(* IEC 61131-3 sources: Test-Git_ESME26/TestProgettoESME_26.fbsproj/AxisModuleLib Migration/AXM_FB_AxisModule.pou.xml.v3^, 40 files *)

(* ---- Additional_active.act.st ---- *)
__METADATA__
{
  "v3Meta": {
    "objectGuid": "95a41eea-732b-4df9-b4b6-dec268632541",
    "objectTypeGuid": "8ac092e5-3128-4e26-9e7e-11016c6684f2",
    "embeddedObjectTypeGuids": [
      "3b83b776-fb25-43b8-99f2-3c507c9143fc"
    ],
    "properties": {},
    "subObjects": {}
  }
}

iq_stAxisModuleItf.stMain.q_etOpMode := AXM_ET_OpMode.Additional;

xAdditionalStart := (xStartFlag OR iq_stAxisModuleItf.stMain.i_xStart) AND NOT stModuleReaction.axReaction[TPL.ET_Reaction.StopEndOfCycle];

iq_stAxisModuleItf.stAdditional.q_xEnable := xAdditionalEnable AND fbDriveEnable.q_xDriveEnabled;
iq_stAxisModuleItf.stAdditional.q_xStart := xAdditionalStart;
iq_stAxisModuleItf.stAdditional.q_xWsSelect := xWsSelect;
iq_stAxisModuleItf.stAdditional.q_xWsStart := xWsStartFlag;

IF iq_stAxisModuleItf.stAdditional.i_etDiag <> GD.ET_Diag.Ok THEN
	stExceptionModuleReaction2.etDiag := GD.ET_Diag.DiagActive;
	stExceptionModuleReaction2.udiDiagExt := AXM_ET_DiagExt.AdditionalModeException;
	stExceptionModuleReaction2.sMsg := SE_CTBX.FC_MultiConcat(	i_sString1 := GD.FC_EtDiagToString(i_etDiag := iq_stAxisModuleItf.stAdditional.i_etDiag),
															i_sString2 := ' ',
															i_sString3 := iq_stAxisModuleItf.stAdditional.i_sDiagExt,
															i_sString4 := SE_CTBX.FC_MultiConcat(	i_sString1 := '(',
																								i_sString2 := UDINT_TO_STRING(iq_stAxisModuleItf.stAdditional.i_udiDiagExt),
																								i_sString3 := ') ',
																								i_sString4 := iq_stAxisModuleItf.stAdditional.i_sMsg));
	ReportException(iq_stException := stExceptionModuleReaction2);
END_IF

xAdditionalActive := iq_stAxisModuleItf.stAdditional.i_xActive;

IF iq_stAxisModuleItf.stAdditional.i_xReady AND NOT iq_stAxisModuleItf.stAdditional.q_xStart THEN
	iq_stAxisModuleItf.stMain.q_etState := AXM_ET_State.AdditionalWaitForStart;
ELSIF iq_stAxisModuleItf.stAdditional.i_xReady AND iq_stAxisModuleItf.stAdditional.q_xStart THEN
	iq_stAxisModuleItf.stMain.q_etState := AXM_ET_State.AdditionalRunning;
ELSE
	IF xAdditionalEnable THEN
		iq_stAxisModuleItf.stMain.q_etState := AXM_ET_State.AdditionalInit;
	ELSE
		iq_stAxisModuleItf.stMain.q_etState := AXM_ET_State.AdditionalExit;
	END_IF
END_IF

(* ---- BrakeRelease_active.act.st ---- *)
__METADATA__
{
  "v3Meta": {
    "objectGuid": "62f6a697-2c31-4fa4-aead-e7013a7e303d",
    "objectTypeGuid": "8ac092e5-3128-4e26-9e7e-11016c6684f2",
    "embeddedObjectTypeGuids": [
      "3b83b776-fb25-43b8-99f2-3c507c9143fc"
    ],
    "properties": {},
    "subObjects": {}
  }
}

iq_stAxisModuleItf.stMain.q_etOpMode := AXM_ET_OpMode.BrakeRelease;

fbBrake(	i_xEnable			:= xBrakeEnable AND NOT fbDriveEnable.q_xDriveEnabled,
			i_xRelease			:= (xStartFlag OR iq_stAxisModuleItf.stMain.i_xStart),
			i_ifDrive			:= iq_stAxisModuleItf.stMain.i_ifDrive,
			q_xActive			=> ,
			q_xReady			=> ,
			q_xReleased			=> iq_stAxisModuleItf.stBrake.q_xBrakeReleased,
			q_etDiag			=> etDiagBuffer,
			q_etDiagExt			=> etDiagExtBufferPDL,
			q_sMsg				=> sDiagMsgBuffer);

DiagTestBrakeRelease(	iq_etDiag		:= fbBrake.q_etDiag,
						iq_etDiagExt	:= fbBrake.q_etDiagExt,
						iq_sMsg			:= fbBrake.q_sMsg);

IF fbBrake.q_xReady AND fbBrake.q_xReleased THEN
	iq_stAxisModuleItf.stMain.q_etState := AXM_ET_State.BrakeReleased;
ELSIF fbBrake.q_xReady AND NOT fbBrake.q_xReleased THEN
	iq_stAxisModuleItf.stMain.q_etState := AXM_ET_State.BrakeClosed;
ELSE
	IF xBrakeEnable THEN
		iq_stAxisModuleItf.stMain.q_etState := AXM_ET_State.BrakeReleaseInit;
	ELSE
		iq_stAxisModuleItf.stMain.q_etState := AXM_ET_State.BrakeReleaseExit;
	END_IF
END_IF

IF NOT xBrakeEnable AND NOT fbBrake.q_xActive THEN
	xBrakeActive := FALSE;
END_IF

(* ---- CancelException.meth.st ---- *)
{attribute 'conditionalshow_all_locals'}
METHOD INTERNAL CancelException
VAR_IN_OUT
	iq_stException	: TPL.ST_Exception;
END_VAR

TPL.FC_SetException(	i_xExceptionActive	:= FALSE,
						iq_stException		:= iq_stException,
						iq_stExceptionList	:= iq_stExceptionList,
						iq_stLogDataList	:= iq_stLogDataList,
						q_etDiag 			=> etDiagBuffer,
						q_etDiagExt 		=> etDiagExtBufferTPL,
						q_sMsg 				=> sDiagMsgBuffer);

(* ---- CheckCmd.meth.st ---- *)
{attribute 'conditionalshow_all_locals'}
METHOD INTERNAL CheckCmd
VAR_INPUT
END_VAR

(*--------------------------------------------------------------------------------------------------*)
(* CheckCMD is checking if CMD is supported by this module *)
(*--------------------------------------------------------------------------------------------------*)
xOpModeCmd:= FALSE;
xCheckCMDError:= FALSE;

IF iq_stStandardModuleItf.iq_diCmd = AXM_ET_Cmd.Homing OR
	iq_stStandardModuleItf.iq_diCmd = AXM_ET_Cmd.Manual OR
	iq_stStandardModuleItf.iq_diCmd = AXM_ET_Cmd.CamCs OR
	iq_stStandardModuleItf.iq_diCmd = AXM_ET_Cmd.CamWs OR
	iq_stStandardModuleItf.iq_diCmd = AXM_ET_Cmd.Endless OR
	iq_stStandardModuleItf.iq_diCmd = AXM_ET_Cmd.Positioning OR
	iq_stStandardModuleItf.iq_diCmd = AXM_ET_Cmd.BrakeRelease OR
	iq_stStandardModuleItf.iq_diCmd = AXM_ET_Cmd.AdditionalCs OR
	iq_stStandardModuleItf.iq_diCmd = AXM_ET_Cmd.AdditionalWs OR
	iq_stStandardModuleItf.iq_diCmd = AXM_ET_Cmd.DriveEnableOff OR
	iq_stStandardModuleItf.iq_diCmd = AXM_ET_Cmd.Stop THEN

	xOpModeCmd := TRUE;

ELSIF  iq_stStandardModuleItf.iq_diCmd = AXM_ET_Cmd.Start OR
		iq_stStandardModuleItf.iq_diCmd = AXM_ET_Cmd.StartTrig OR
		iq_stStandardModuleItf.iq_diCmd = AXM_ET_Cmd.StartTrigWaitInPos OR
		iq_stStandardModuleItf.iq_diCmd = AXM_ET_Cmd.Hold OR
		iq_stStandardModuleItf.iq_diCmd = AXM_ET_Cmd.WsStart OR
		iq_stStandardModuleItf.iq_diCmd = AXM_ET_Cmd.DriveEnableOn THEN

		xOpModeCmd:= FALSE;
ELSE
	xCheckCMDError := TRUE;
END_IF

(* ---- CmdControl_active.act.st ---- *)
__METADATA__
{
  "v3Meta": {
    "objectGuid": "07d6aa58-0565-4f47-8048-7bdd25741778",
    "objectTypeGuid": "8ac092e5-3128-4e26-9e7e-11016c6684f2",
    "embeddedObjectTypeGuids": [
      "3b83b776-fb25-43b8-99f2-3c507c9143fc"
    ],
    "properties": {},
    "subObjects": {}
  }
}

(* CMD execution

	algorithm:
	----------

	detect new command?
		check command?
			execute command;
		end
	end

	is command running (at least one cycle)?
		is command finished?
			signal success/unsuccessful
		end
	end
*)

xCommandAcceptedInThisCycle := FALSE;

(* Detect new command *)
IF(iq_stStandardModuleItf.i_xEnable) THEN
	IF (iq_stStandardModuleItf.iq_diCmd > 0 AND (NOT iq_stStandardModuleItf.q_xCmdActive (* In case no command is active *)
			OR iq_stStandardModuleItf.iq_diCmd <> iq_stStandardModuleItf.q_diCmdActive) (* In case a command is active *)) THEN

		xCommandRefused := FALSE; (* Flag is set by RefuseCommand() action *)

(****** Check if command execution is possible ******)
		CheckCMD();
		IF(xCheckCMDError) THEN
			(*** Check for unknown command ***)
			stExceptionCmdUnknown.sMsg := Standard.CONCAT('Cmd unknown: ',DINT_TO_STRING(iq_stStandardModuleItf.iq_diCmd));
			ReportException(iq_stException := stExceptionCmdUnknown);
			RefuseCommand();
		ELSE
			(*** Check for impossible overwrite ***)
			IF(iq_stStandardModuleItf.q_xCmdActive AND NOT((iq_stStandardModuleItf.iq_diCmd = AXM_ET_Cmd.Stop) OR
															(iq_stStandardModuleItf.iq_diCmd = AXM_ET_Cmd.BrakeRelease) OR
															((iq_stStandardModuleItf.iq_diCmd = AXM_ET_Cmd.Hold) AND (iq_stAxisModuleItf.stMain.q_etOpMode = AXM_ET_OpMode.Positioning) AND (iq_stStandardModuleItf.q_diCmdActive = AXM_ET_Cmd.Start)) OR
															((iq_stStandardModuleItf.iq_diCmd = AXM_ET_Cmd.Start) AND (iq_stAxisModuleItf.stMain.q_etOpMode = AXM_ET_OpMode.Endless) AND (iq_stStandardModuleItf.q_diCmdActive = AXM_ET_Cmd.Hold)))) THEN
				stExceptionCmdImpossibleOverwrite.sMsg := SE_CTBX.FC_MultiConcat(	i_sString1 := 'Cmd impossible: ',
																				//i_sString2 := iq_stStandardModuleItf.iq_diCmd
																				i_sString2 := AXM_FC_EtCmdToString(i_etCmd := iq_stStandardModuleItf.iq_diCmd),
																				i_sString3 := '; Cmd active: ',
																				i_sString4 := AXM_FC_EtCmdToString(i_etCmd := iq_stStandardModuleItf.q_diCmdActive) );
				ReportException(iq_stException := stExceptionCmdImpossibleOverwrite);
				RefuseCommand();
			ELSE
				(*** Check for impossible state ***)
				IF (((iq_stAxisModuleItf.stMain.q_etState = AXM_ET_State.NoOpDriveDisabled) OR (iq_stAxisModuleItf.stMain.q_etState = AXM_ET_State.NoOpDriveEnabled) ) AND
																								((iq_stStandardModuleItf.iq_diCmd = AXM_ET_Cmd.Start) OR
																								(iq_stStandardModuleItf.iq_diCmd = AXM_ET_Cmd.WsStart) OR
																								(iq_stStandardModuleItf.iq_diCmd = AXM_ET_Cmd.StartTrig) OR
																								(iq_stStandardModuleItf.iq_diCmd = AXM_ET_Cmd.StartTrigWaitInPos)) ) OR
					((iq_stAxisModuleItf.stMain.q_etState <> AXM_ET_State.MultiCamWaitForWsStart) AND (iq_stAxisModuleItf.stMain.q_etState <> AXM_ET_State.MultiCamRunning) AND (iq_stAxisModuleItf.stMain.q_etOpMode <> AXM_ET_OpMode.Additional) AND (iq_stStandardModuleItf.iq_diCmd = AXM_ET_Cmd.WsStart)) OR
					((iq_stAxisModuleItf.stMain.q_etState = AXM_ET_State.MultiCamWaitForWsStart) AND ((iq_stStandardModuleItf.iq_diCmd = AXM_ET_Cmd.WsStart) AND ((iq_stAxisModuleItf.stMultiCam.i_etWsMode = PDL_ET_MultiCamWsMode.StoredCamShowCamPosition) OR
																																		(iq_stAxisModuleItf.stMultiCam.i_etWsMode = PDL_ET_MultiCamWsMode.NewCamShowCamPosition)) ) ) OR
					((iq_stAxisModuleItf.stMain.q_etOpMode = AXM_ET_OpMode.Manual) AND ((iq_stStandardModuleItf.iq_diCmd = AXM_ET_Cmd.Hold) OR
																											(iq_stStandardModuleItf.iq_diCmd = AXM_ET_Cmd.Start)) ) OR
					((iq_stAxisModuleItf.stMain.q_etOpMode <> AXM_ET_OpMode.Positioning) AND (iq_stStandardModuleItf.iq_diCmd = AXM_ET_Cmd.StartTrigWaitInPos)) OR
					((iq_stAxisModuleItf.stMain.q_etOpMode <> AXM_ET_OpMode.Endless) AND (iq_stAxisModuleItf.stMain.q_etOpMode <> AXM_ET_OpMode.MultiCam) AND (iq_stAxisModuleItf.stMain.q_etOpMode <> AXM_ET_OpMode.Positioning) AND (iq_stStandardModuleItf.iq_diCmd = AXM_ET_Cmd.StartTrig))
					THEN
					stExceptionCmdImpossibleState.sMsg := SE_CTBX.FC_MultiConcat(	i_sString1 := 'Cmd impossible: ',
																				i_sString2 := AXM_FC_EtCmdToString(i_etCmd := iq_stStandardModuleItf.iq_diCmd),
																				i_sString3 := '; State: ',
																				i_sString4 := AXM_FC_EtStateToString(i_etState := iq_stAxisModuleItf.stMain.q_etState) );
					ReportException(iq_stException := stExceptionCmdImpossibleState);
					RefuseCommand();
				ELSIF ((iq_stAxisModuleItf.stMain.q_etOpMode = AXM_ET_OpMode.Homing OR
						iq_stAxisModuleItf.stMain.q_etOpMode = AXM_ET_OpMode.Manual OR
						iq_stAxisModuleItf.stMain.q_etOpMode = AXM_ET_OpMode.MultiCam OR
						iq_stAxisModuleItf.stMain.q_etOpMode = AXM_ET_OpMode.Endless OR
						iq_stAxisModuleItf.stMain.q_etOpMode = AXM_ET_OpMode.Positioning OR
						iq_stAxisModuleItf.stMain.q_etOpMode = AXM_ET_OpMode.BrakeRelease OR
						iq_stAxisModuleItf.stMain.q_etOpMode = AXM_ET_OpMode.Additional) AND ((iq_stAxisModuleItf.stMain.i_xStart OR xStartBitLastCycle) AND (iq_stStandardModuleItf.iq_diCMD = AXM_ET_Cmd.Start OR
																																						iq_stStandardModuleItf.iq_diCMD = AXM_ET_Cmd.Hold OR
																																						iq_stStandardModuleItf.iq_diCMD = AXM_ET_Cmd.StartTrig OR
																																						iq_stStandardModuleItf.iq_diCMD = AXM_ET_Cmd.StartTrigWaitInPos) )) THEN
					IF(iq_stAxisModuleItf.stMain.i_xStart) THEN
						stExceptionCmdImpossibleState.sMsg := SE_CTBX.FC_MultiConcat(	i_sString1 := 'Cmd impossible: ',
																					i_sString2 := AXM_FC_EtCmdToString(i_etCmd := iq_stStandardModuleItf.iq_diCmd),
																					i_sString3 := '; State: ',
																					i_sString4 := 'xStart input is TRUE');
						ReportException(iq_stException := stExceptionCmdImpossibleState);
						RefuseCommand();
					ELSE
						stExceptionCmdImpossibleState.sMsg := SE_CTBX.FC_MultiConcat(	i_sString1 := 'Cmd impossible: ',
																					i_sString2 := AXM_FC_EtCmdToString(i_etCmd := iq_stStandardModuleItf.iq_diCmd),
																					i_sString3 := '; State: ',
																					i_sString4 := 'xStart input was TRUE last cycle');
						ReportException(iq_stException := stExceptionCmdImpossibleState);
						RefuseCommand();
					END_IF
				ELSE
					(*** Check for impossible commands due to active error reactions ***)
					IF (stModuleReaction.axReaction[TPL.ET_Reaction.AsyncStop]
						OR stModuleReaction.axReaction[TPL.ET_Reaction.SyncStopEH]
						OR stModuleReaction.axReaction[TPL.ET_Reaction.SyncStopEL]
						OR stModuleReaction.axReaction[TPL.ET_Reaction.StopEndOfCycle])
						AND NOT (iq_stAxisModuleItf.stMain.q_etOpMode = AXM_ET_OpMode.BrakeRelease)
						AND	((iq_stStandardModuleItf.iq_diCmd = AXM_ET_Cmd.Start) OR
							(iq_stStandardModuleItf.iq_diCmd = AXM_ET_Cmd.WsStart) OR
							(iq_stStandardModuleItf.iq_diCmd = AXM_ET_Cmd.StartTrig) OR
							(iq_stStandardModuleItf.iq_diCmd = AXM_ET_Cmd.StartTrigWaitInPos)) THEN (* Start impossible if error reaction 4 or higher *)
							stWarningCmdImpossibleReaction.sMsg := SE_CTBX.FC_MultiConcat(	i_sString1 := 'Cmd impossible: ',
																						i_sString2 := AXM_FC_EtCmdToString(i_etCmd := iq_stStandardModuleItf.iq_diCmd),
																						i_sString3 := '; Reaction: ',
																						i_sString4 := TPL.FC_GetStandardReactionName(iq_stReaction := stModuleReaction));
							ReportException(iq_stException := stWarningCmdImpossibleReaction);
							RefuseCommand();
					ELSIF ((stModuleReaction.axReaction[TPL.ET_Reaction.AsyncStop]
							OR stModuleReaction.axReaction[TPL.ET_Reaction.SyncStopEH]
							OR stModuleReaction.axReaction[TPL.ET_Reaction.SyncStopEL] )
							AND xOpModeCmd AND
							NOT ((iq_stStandardModuleItf.iq_diCmd = AXM_ET_Cmd.Stop) OR (iq_stStandardModuleItf.iq_diCmd = AXM_ET_Cmd.DriveEnableOff) OR (iq_stStandardModuleItf.iq_diCmd = AXM_ET_Cmd.BrakeRelease)) ) THEN
							stWarningCmdImpossibleReaction.sMsg := SE_CTBX.FC_MultiConcat(	i_sString1 := 'Cmd impossible: ',
																						i_sString2 := AXM_FC_EtCmdToString(i_etCmd := iq_stStandardModuleItf.iq_diCmd),
																						i_sString3 := '; Reaction: ',
																						i_sString4 := TPL.FC_GetStandardReactionName(iq_stReaction := stModuleReaction));
							ReportException(iq_stException := stWarningCmdImpossibleReaction);
							RefuseCommand();
					ELSIF ((stModuleReaction.axReaction[TPL.ET_Reaction.AsyncStop]
							OR stModuleReaction.axReaction[TPL.ET_Reaction.SyncStopEL])
							AND (iq_stStandardModuleItf.iq_diCmd = AXM_ET_Cmd.DriveEnableOn)) THEN
							stWarningCmdImpossibleReaction.sMsg := SE_CTBX.FC_MultiConcat(	i_sString1 := 'Cmd impossible: ',
																						i_sString2 := AXM_FC_EtCmdToString(i_etCmd := iq_stStandardModuleItf.iq_diCmd),
																						i_sString3 := '; Reaction: ',
																						i_sString4 := TPL.FC_GetStandardReactionName(iq_stReaction := stModuleReaction));
							ReportException(iq_stException := stWarningCmdImpossibleReaction);
							RefuseCommand();
					END_IF
				END_IF
			END_IF
		END_IF

		IF(NOT xCommandRefused) THEN (* Command has passed all checks, execute command *)
			(* Accept command *)
			iq_stStandardModuleItf.q_xCmdActive := TRUE;
			iq_stStandardModuleItf.q_xCmdDone := FALSE;
			iq_stStandardModuleItf.q_diCmdActive := iq_stStandardModuleItf.iq_diCmd;

			xCommandAcceptedInThisCycle := TRUE; (* Signal for command done checks *)
			IF fbLoggerPoint.etLogLevel >= APL.ET_LogLevel.UserAction THEN
				fbLoggerPoint.AddLogEntry(	i_etLogLevel	:= APL.ET_LogLevel.UserAction,
											i_etDiag		:= GD.ET_Diag.Ok,
											i_udiDiagExt	:= AXM_ET_DiagExt.Ok,
											i_sMessage		:= Standard.CONCAT(Standard.CONCAT(Standard.CONCAT('Command executing: ', AXM_FC_EtCmdToString(i_etCmd := iq_stStandardModuleItf.iq_diCmd)),' number: '),DINT_TO_STRING(iq_stStandardModuleItf.iq_diCmd)),
											q_etDiag		:= ,
											q_etDiagExt		:= );
			END_IF

			IF(xOpModeCmd) THEN
				DisableAllJobs();
				xWsSelect			:= FALSE;
				xWsStartFlag		:= FALSE;

				CASE iq_stStandardModuleItf.iq_diCmd OF
				AXM_ET_Cmd.Stop:
					(* Do nothing, disabled OpMode flags automatically lead to NoOp *)
					xStartFlag := FALSE;

				AXM_ET_Cmd.Homing:
					xRefEnable := TRUE;

					IF iq_stAxisModuleItf.stHome.stSetPos.i_xKeepPowerDisabled AND
						( iq_stAxisModuleItf.stHome.i_etMode = PDL_ET_HomeMode.RestorePosFromAxisEncoder
						OR iq_stAxisModuleItf.stHome.i_etMode = PDL_ET_HomeMode.RestorePosFromRetain
						OR iq_stAxisModuleItf.stHome.i_etMode = PDL_ET_HomeMode.SetPosAxisAndLogEncoderPosition
						OR iq_stAxisModuleItf.stHome.i_etMode = PDL_ET_HomeMode.SetPosAxisPosition
						OR iq_stAxisModuleItf.stHome.i_etMode = PDL_ET_HomeMode.SetPosLogEncoderPosition )THEN
						xCMDPowerOn := FALSE;
					ELSE
						xCMDPowerOn := TRUE;
					END_IF

					IF NOT (iq_stAxisModuleItf.stMain.q_etOpMode = AXM_ET_OpMode.Homing) THEN
						xStartFlag := FALSE;
					END_IF

				AXM_ET_Cmd.Manual:
					xManEnable := TRUE;
					xCMDPowerOn := TRUE;

				AXM_ET_Cmd.CamCs:
					xCamEnable := TRUE;
					xCMDPowerOn := TRUE;
					xWsSelect := FALSE;
					xWsStartFlag := FALSE;
					IF NOT (iq_stAxisModuleItf.stMain.q_etOpMode = AXM_ET_OpMode.MultiCam) THEN
						xStartFlag := FALSE;
					END_IF

				AXM_ET_Cmd.CamWs:
					xCamEnable := TRUE;
					xCMDPowerOn := TRUE;
					xWsSelect := TRUE;
					xWsStartFlag := FALSE;
					IF NOT (iq_stAxisModuleItf.stMain.q_etOpMode = AXM_ET_OpMode.MultiCam) THEN
						xStartFlag := FALSE;
					END_IF

				AXM_ET_Cmd.Endless:
					xEndlessEnable := TRUE;
					xCMDPowerOn := TRUE;
					IF NOT (iq_stAxisModuleItf.stMain.q_etOpMode = AXM_ET_OpMode.Endless) THEN
						xStartFlag := FALSE;
					END_IF

				AXM_ET_Cmd.Positioning:
					xPosEnable := TRUE;
					xCMDPowerOn := TRUE;
					IF NOT (iq_stAxisModuleItf.stMain.q_etOpMode = AXM_ET_OpMode.Positioning) THEN
						xStartFlag := FALSE;
					END_IF

				AXM_ET_Cmd.BrakeRelease:
					xBrakeEnable := TRUE;
					xCMDPowerOn := FALSE;
					IF NOT (iq_stAxisModuleItf.stMain.q_etOpMode = AXM_ET_OpMode.BrakeRelease) THEN
						xStartFlag := FALSE;
					END_IF

				AXM_ET_Cmd.AdditionalCs:
					xAdditionalEnable := TRUE;
					xCMDPowerOn := TRUE;
					xWsSelect := FALSE;
					xWsStartFlag := FALSE;
					IF NOT (iq_stAxisModuleItf.stMain.q_etOpMode = AXM_ET_OpMode.Additional) THEN
						xStartFlag := FALSE;
					END_IF

				AXM_ET_Cmd.AdditionalWs:
					xAdditionalEnable := TRUE;
					xCMDPowerOn := TRUE;
					xWsSelect := TRUE;
					xWsStartFlag := FALSE;
					IF NOT (iq_stAxisModuleItf.stMain.q_etOpMode = AXM_ET_OpMode.Additional) THEN
						xStartFlag := FALSE;
					END_IF

				AXM_ET_Cmd.DriveEnableOff:
					xCMDPowerOn := FALSE;
					xStartFlag := FALSE;
				ELSE
					stExceptionModuleReaction1.etDiag := GD.ET_Diag.UnexpectedProgramBehavior;
					stExceptionModuleReaction1.udiDiagExt := AXM_ET_DiagExt.UnknownCase;
					stExceptionModuleReaction1.sMsg := '';
					ReportException(iq_stException := stExceptionModuleReaction1);
				END_CASE
			ELSE
				CASE iq_stStandardModuleItf.iq_diCmd OF
				AXM_ET_Cmd.Start:
					xStartFlag := TRUE;
					IF (iq_stAxisModuleItf.stMain.q_etOpMode = AXM_ET_OpMode.Homing) THEN
						(* Reset HomeOk when a new homing is started *)
						iq_stAxisModuleItf.stMain.q_xHomeOk := FALSE;
					END_IF

				AXM_ET_Cmd.StartTrig:
					xStartFlag := TRUE;

				AXM_ET_Cmd.StartTrigWaitInPos:
					xStartFlag := TRUE;

				AXM_ET_Cmd.WsStart:
					xWsStartFlag := TRUE;
					(* In additional mode it has to be possible to set WsStart independent of start *)
					IF NOT (iq_stAxisModuleItf.stMain.q_etOpMode = AXM_ET_OpMode.Additional) THEN
						xStartFlag  := TRUE;
					END_IF

				AXM_ET_Cmd.Hold:
					xStartFlag := FALSE;

				AXM_ET_Cmd.DriveEnableOn:
					xCMDPowerOn := TRUE;

				ELSE
					stExceptionModuleReaction1.etDiag := GD.ET_Diag.UnexpectedProgramBehavior;
					stExceptionModuleReaction1.udiDiagExt := AXM_ET_DiagExt.UnknownCase;
					stExceptionModuleReaction1.sMsg := '';
					ReportException(iq_stException := stExceptionModuleReaction1);
				END_CASE

			END_IF
		END_IF (* New command? *)
	END_IF

(********************************************* Check successful and unsucessful of given commands ****************************************)

	(* Check if active command is done or is stopped by an error *)
	IF(NOT xCommandAcceptedInThisCycle) THEN (* Don't execute these checks if we accepted a new command in this cycle
		to ensure that execution of every command requires a minimum of 2 cycles *)

		IF(iq_stStandardModuleItf.q_xCmdActive) THEN
			CASE iq_stStandardModuleItf.iq_diCmd OF
			AXM_ET_Cmd.Homing:
				(* Successful *)
				IF (iq_stAxisModuleItf.stMain.q_etOpMode = AXM_ET_OpMode.Homing) AND NOT (iq_stAxisModuleItf.stMain.q_etState = AXM_ET_State.HomingInit) THEN
					SignalSuccessfulExecution();
				END_IF
				(* Unsucessful *)
				IF(stModuleReaction.axReaction[TPL.ET_Reaction.AsyncStop]
					OR stModuleReaction.axReaction[TPL.ET_Reaction.SyncStopEH]
					OR stModuleReaction.axReaction[TPL.ET_Reaction.SyncStopEL]) THEN
					SignalUnsuccessfulExecution();
				END_IF

			AXM_ET_Cmd.Manual:
				(* Successful *)
				IF (iq_stAxisModuleItf.stMain.q_etOpMode = AXM_ET_OpMode.Manual) AND NOT (iq_stAxisModuleItf.stMain.q_etState = AXM_ET_State.ManualInit) THEN
					SignalSuccessfulExecution();
				END_IF
				(* Unsucessful *)
				IF(stModuleReaction.axReaction[TPL.ET_Reaction.AsyncStop]
					OR stModuleReaction.axReaction[TPL.ET_Reaction.SyncStopEH]
					OR stModuleReaction.axReaction[TPL.ET_Reaction.SyncStopEL]) THEN
					SignalUnsuccessfulExecution();
				END_IF

			AXM_ET_Cmd.CamCs:
				(* Successful *)
				IF (iq_stAxisModuleItf.stMain.q_etOpMode = AXM_ET_OpMode.MultiCam) AND NOT (iq_stAxisModuleItf.stMain.q_etState = AXM_ET_State.MultiCamInit) THEN
					SignalSuccessfulExecution();
				END_IF
				(* Unsucessful *)
				IF(stModuleReaction.axReaction[TPL.ET_Reaction.AsyncStop]
					OR stModuleReaction.axReaction[TPL.ET_Reaction.SyncStopEH]
					OR stModuleReaction.axReaction[TPL.ET_Reaction.SyncStopEL]) THEN
					SignalUnsuccessfulExecution();
				END_IF

			AXM_ET_Cmd.CamWs:
				(* Successful *)
				IF (iq_stAxisModuleItf.stMain.q_etOpMode = AXM_ET_OpMode.MultiCam) AND NOT (iq_stAxisModuleItf.stMain.q_etState = AXM_ET_State.MultiCamInit) THEN
					SignalSuccessfulExecution();
				END_IF
				(* Unsucessful *)
				IF(stModuleReaction.axReaction[TPL.ET_Reaction.AsyncStop]
					OR stModuleReaction.axReaction[TPL.ET_Reaction.SyncStopEH]
					OR stModuleReaction.axReaction[TPL.ET_Reaction.SyncStopEL]) THEN
					SignalUnsuccessfulExecution();
				END_IF

			AXM_ET_Cmd.Endless:
				(* Successful *)
				IF (iq_stAxisModuleItf.stMain.q_etOpMode = AXM_ET_OpMode.Endless) AND NOT (iq_stAxisModuleItf.stMain.q_etState = AXM_ET_State.EndlessInit) THEN
					SignalSuccessfulExecution();
				END_IF
				(* Unsucessful *)
				IF(stModuleReaction.axReaction[TPL.ET_Reaction.AsyncStop]
					OR stModuleReaction.axReaction[TPL.ET_Reaction.SyncStopEH]
					OR stModuleReaction.axReaction[TPL.ET_Reaction.SyncStopEL]) THEN
					SignalUnsuccessfulExecution();
				END_IF

			AXM_ET_Cmd.Positioning:
				(* Successful *)
				IF (iq_stAxisModuleItf.stMain.q_etOpMode = AXM_ET_OpMode.Positioning) AND NOT (iq_stAxisModuleItf.stMain.q_etState = AXM_ET_State.PositioningInit) THEN
					SignalSuccessfulExecution();
				END_IF
				(* Unsucessful *)
				IF(stModuleReaction.axReaction[TPL.ET_Reaction.AsyncStop]
					OR stModuleReaction.axReaction[TPL.ET_Reaction.SyncStopEH]
					OR stModuleReaction.axReaction[TPL.ET_Reaction.SyncStopEL]) THEN
					SignalUnsuccessfulExecution();
				END_IF

			AXM_ET_Cmd.BrakeRelease:
				(* Successful *)
				IF (iq_stAxisModuleItf.stMain.q_etOpMode = AXM_ET_OpMode.BrakeRelease) AND
					( (NOT fbBrake.i_xRelease AND (iq_stAxisModuleItf.stMain.q_etState = AXM_ET_State.BrakeClosed)) OR
					(fbBrake.i_xRelease AND (iq_stAxisModuleItf.stMain.q_etState = AXM_ET_State.BrakeReleased)) ) THEN
					// real axis can still be in state brake open if gone to brake release opmode,
					// therefore delay signal cmd successfull till brake closed is reached
					SignalSuccessfulExecution();
				END_IF

			AXM_ET_Cmd.AdditionalCs:
				(* Successful *)
				IF (iq_stAxisModuleItf.stMain.q_etOpMode = AXM_ET_OpMode.Additional) AND NOT (iq_stAxisModuleItf.stMain.q_etState = AXM_ET_State.AdditionalInit) THEN
					SignalSuccessfulExecution();
				END_IF
				(* Unsucessful *)
				IF(stModuleReaction.axReaction[TPL.ET_Reaction.AsyncStop]
					OR stModuleReaction.axReaction[TPL.ET_Reaction.SyncStopEH]
					OR stModuleReaction.axReaction[TPL.ET_Reaction.SyncStopEL]) THEN
					SignalUnsuccessfulExecution();
				END_IF

			AXM_ET_Cmd.AdditionalWs:
				(* Successful *)
				IF (iq_stAxisModuleItf.stMain.q_etOpMode = AXM_ET_OpMode.Additional) AND NOT (iq_stAxisModuleItf.stMain.q_etState = AXM_ET_State.AdditionalInit) THEN
					SignalSuccessfulExecution();
				END_IF
				(* Unsucessful *)
				IF(stModuleReaction.axReaction[TPL.ET_Reaction.AsyncStop]
					OR stModuleReaction.axReaction[TPL.ET_Reaction.SyncStopEH]
					OR stModuleReaction.axReaction[TPL.ET_Reaction.SyncStopEL]) THEN
					SignalUnsuccessfulExecution();
				END_IF

			AXM_ET_Cmd.Start:
				(* Successful *)
				IF ((iq_stAxisModuleItf.stMain.q_etState = AXM_ET_State.HomingWaitForStart) AND iq_stAxisModuleItf.stMain.q_xHomeOk) OR
					(iq_stAxisModuleItf.stMain.q_etState = AXM_ET_State.HomingDone) OR
					(iq_stAxisModuleItf.stMain.q_etState = AXM_ET_State.MultiCamWaitForWsStart) OR
					(iq_stAxisModuleItf.stMain.q_etState = AXM_ET_State.MultiCamRunning) OR
					(iq_stAxisModuleItf.stMain.q_etState = AXM_ET_State.EndlessRunning) OR
					(iq_stAxisModuleItf.stMain.q_etState = AXM_ET_State.PositioningRunning) OR
					(iq_stAxisModuleItf.stMain.q_etState = AXM_ET_State.BrakeReleased) OR
					((iq_stAxisModuleItf.stMain.q_etOpMode = AXM_ET_OpMode.Additional) AND iq_stAxisModuleItf.stAdditional.i_xActionCmdDone) THEN
					SignalSuccessfulExecution();
				END_IF
				(* Unsucesful *)
				IF(stModuleReaction.axReaction[TPL.ET_Reaction.AsyncStop]
					OR stModuleReaction.axReaction[TPL.ET_Reaction.SyncStopEH]
					OR stModuleReaction.axReaction[TPL.ET_Reaction.SyncStopEL]
					OR stModuleReaction.axReaction[TPL.ET_Reaction.StopEndOfCycle])
					AND NOT (iq_stAxisModuleItf.stMain.q_etOpMode = AXM_ET_OpMode.BrakeRelease) THEN
					SignalUnsuccessfulExecution();
				END_IF

			AXM_ET_Cmd.StartTrig:
				(* Successful *)
				IF (iq_stAxisModuleItf.stMain.q_etState = AXM_ET_State.PositioningRunning) OR
					(iq_stAxisModuleItf.stMain.q_etState = AXM_ET_State.MultiCamRunning) OR
					(iq_stAxisModuleItf.stMain.q_etState = AXM_ET_State.EndlessRunning) THEN
					xStartFlag := FALSE;
					SignalSuccessfulExecution();
				END_IF
				(* Unsucesful *)
				IF(stModuleReaction.axReaction[TPL.ET_Reaction.AsyncStop]
					OR stModuleReaction.axReaction[TPL.ET_Reaction.SyncStopEH]
					OR stModuleReaction.axReaction[TPL.ET_Reaction.SyncStopEL]
					)
					AND NOT (iq_stAxisModuleItf.stMain.q_etOpMode = AXM_ET_OpMode.BrakeRelease) THEN
					SignalUnsuccessfulExecution();
				END_IF

			AXM_ET_Cmd.StartTrigWaitInPos:
				(* Successful *)
				IF fbVarioPos.q_xInPosition THEN
					xStartFlag := FALSE;
					SignalSuccessfulExecution();
				END_IF
				(* Unsucesful *)
				IF(stModuleReaction.axReaction[TPL.ET_Reaction.AsyncStop]
					OR stModuleReaction.axReaction[TPL.ET_Reaction.SyncStopEH]
					OR stModuleReaction.axReaction[TPL.ET_Reaction.SyncStopEL]
					)
					AND NOT (iq_stAxisModuleItf.stMain.q_etOpMode = AXM_ET_OpMode.BrakeRelease) THEN
					SignalUnsuccessfulExecution();
				END_IF

			AXM_ET_Cmd.Stop:
				(* Successful *)
				IF (iq_stAxisModuleItf.stMain.q_etState = AXM_ET_State.NoOpDriveDisabled) OR
					(iq_stAxisModuleItf.stMain.q_etState = AXM_ET_State.NoOpDriveEnabled) THEN
					iq_stAxisModuleItf.stMain.q_etOpMode := AXM_ET_OpMode.NoOp;
					SignalSuccessfulExecution();
				END_IF

			AXM_ET_Cmd.Hold:
				IF iq_stAxisModuleItf.stMain.i_xStart THEN
					stExceptionModuleReaction2.sMsg := 'rising edge of xStart input during execution of CMD Hold';
					ReportException(iq_stException := stExceptionModuleReaction2);
					RefuseCommand();
				ELSIF (* Successful *)
					(iq_stAxisModuleItf.stMain.q_etState = AXM_ET_State.HomingWaitForStart) OR
					(iq_stAxisModuleItf.stMain.q_etState = AXM_ET_State.MultiCamWaitForStart) OR
					(iq_stAxisModuleItf.stMain.q_etState = AXM_ET_State.EndlessWaitForStart) OR
					(iq_stAxisModuleItf.stMain.q_etState = AXM_ET_State.PositioningWaitForStart) OR
					(iq_stAxisModuleItf.stMain.q_etState = AXM_ET_State.BrakeClosed) OR
					(iq_stAxisModuleItf.stMain.q_etState = AXM_ET_State.AdditionalWaitForStart) OR
					(iq_stAxisModuleItf.stMain.q_etState = AXM_ET_State.NoOpDriveDisabled) OR
					(iq_stAxisModuleItf.stMain.q_etState = AXM_ET_State.NoOpDriveEnabled) OR
					((iq_stAxisModuleItf.stMain.q_etOpMode = AXM_ET_OpMode.Additional) AND iq_stAxisModuleItf.stAdditional.i_xActionCmdDone) THEN
					SignalSuccessfulExecution();
				ELSIF (* Unsucessful *)
					(stModuleReaction.axReaction[TPL.ET_Reaction.AsyncStop]
					OR stModuleReaction.axReaction[TPL.ET_Reaction.SyncStopEH]
					OR stModuleReaction.axReaction[TPL.ET_Reaction.SyncStopEL]) AND NOT (iq_stAxisModuleItf.stMain.q_etOpMode = AXM_ET_OpMode.BrakeRelease) THEN
					SignalUnsuccessfulExecution();
				END_IF

			AXM_ET_Cmd.WsStart:
				(* Successful *)
				IF ((iq_stAxisModuleItf.stMain.q_etState = AXM_ET_State.HomingWaitForStart) AND iq_stAxisModuleItf.stMain.q_xHomeOk) OR
					(iq_stAxisModuleItf.stMain.q_etState = AXM_ET_State.MultiCamRunning) OR
					(iq_stAxisModuleItf.stMain.q_etState = AXM_ET_State.EndlessRunning) OR
					(iq_stAxisModuleItf.stMain.q_etState = AXM_ET_State.PositioningRunning) OR
					(iq_stAxisModuleItf.stMain.q_etState = AXM_ET_State.BrakeReleased) OR
					((iq_stAxisModuleItf.stMain.q_etOpMode = AXM_ET_OpMode.Additional) AND iq_stAxisModuleItf.stAdditional.i_xActionCmdDone) THEN
					SignalSuccessfulExecution();
				END_IF
				(* Unsucesful *)
				IF(stModuleReaction.axReaction[TPL.ET_Reaction.AsyncStop]
					OR stModuleReaction.axReaction[TPL.ET_Reaction.SyncStopEH]
					OR stModuleReaction.axReaction[TPL.ET_Reaction.SyncStopEL]
					OR stModuleReaction.axReaction[TPL.ET_Reaction.StopEndOfCycle]) THEN
					SignalUnsuccessfulExecution();
				END_IF

			AXM_ET_Cmd.DriveEnableOn:
				(* Successful *)
				IF(etPowerState = AXM_ET_PowerState.PowerOn) THEN
					SignalSuccessfulExecution();
				END_IF
				(* Unsucessful *)
				IF(stModuleReaction.axReaction[TPL.ET_Reaction.AsyncStop]
					OR stModuleReaction.axReaction[TPL.ET_Reaction.SyncStopEH]
					OR stModuleReaction.axReaction[TPL.ET_Reaction.SyncStopEL]) THEN
					SignalUnsuccessfulExecution();
				END_IF

			AXM_ET_Cmd.DriveEnableOff:
				(* Successful *)
				IF(etPowerState = AXM_ET_PowerState.PowerOff) THEN
					SignalSuccessfulExecution();
				END_IF

			ELSE
				stExceptionModuleReaction1.etDiag := GD.ET_Diag.UnexpectedProgramBehavior;
				stExceptionModuleReaction1.udiDiagExt := AXM_ET_DiagExt.UnknownCase;
				stExceptionModuleReaction1.sMsg := '';
				ReportException(iq_stException := stExceptionModuleReaction1);
			END_CASE
		END_IF
	END_IF
ELSE
	(* Module is going to be disabled *)
	IF xEnableFlag THEN
		etPowerState := AXM_ET_PowerState.WaitForDisabled;
		IF fbLoggerPoint.etLogLevel >= APL.ET_LogLevel.UserAction THEN
			fbLoggerPoint.AddLogEntry(	i_etLogLevel	:= APL.ET_LogLevel.UserAction,
										i_etDiag		:= GD.ET_Diag.Ok,
										i_udiDiagExt	:= AXM_ET_DiagExt.Ok,
										i_sMessage		:= 'disabeling Module',
										q_etDiag		:= ,
										q_etDiagExt		:= );
		END_IF
	END_IF
	iq_stStandardModuleItf.q_xReady := FALSE;
	xEnableFlag := FALSE;
	xCMDPowerOn := FALSE;
	DisableAllJobs();
	xStartFlag := FALSE;
	xWsSelect := FALSE;
	xWsStartFlag := FALSE;
	IF(iq_stStandardModuleItf.q_xCmdActive) THEN (* If a command is currently active, cancel its execution *)
		SignalUnsuccessfulExecution();
	ELSE
		InactiveCmdExecution(); (* Command processing as if we were disabled *)
	END_IF
END_IF
xStartBitLastCycle := iq_stAxisModuleItf.stMain.i_xStart;

(* ---- DiagQuit.meth.st ---- *)
{attribute 'conditionalshow_all_locals'}
METHOD INTERNAL DiagQuit
VAR_INPUT
END_VAR

IF(iq_stStandardModuleItf.i_xDiagQuit AND NOT xDiagQuitFlag) THEN
	(* Rising edge of error quit *)
	xDiagQuitFlag := TRUE;
	xNotAbleToSetException := FALSE;
	iq_stStandardModuleItf.q_xException := FALSE;

	FOR udii := 1 TO TPL.ET_Reaction.MainsContactorOff DO
		stLocalReaction.axReaction[udii] := FALSE;
	END_FOR

	IF(iq_stStandardModuleItf.iq_diCMD < 0) THEN
		iq_stStandardModuleItf.iq_diCMD := 0;
	END_IF
	IF fbLoggerPoint.etLogLevel >= APL.ET_LogLevel.UserAction THEN
		fbLoggerPoint.AddLogEntry(	i_etLogLevel	:= APL.ET_LogLevel.UserAction,
									i_etDiag		:= GD.ET_Diag.Ok,
									i_udiDiagExt	:= AXM_ET_DiagExt.Ok,
									i_sMessage		:= 'Diag Quit',
									q_etDiag		:= ,
									q_etDiagExt		:= );
	END_IF
ELSIF(NOT iq_stStandardModuleItf.i_xDiagQuit AND xDiagQuitFlag) THEN
	xDiagQuitFlag := FALSE;
END_IF

(* ---- DiagTestBrakeRelease.meth.st ---- *)
{attribute 'conditionalshow_all_locals'}
METHOD INTERNAL DiagTestBrakeRelease
VAR_IN_OUT
	iq_etDiag		: GD.ET_Diag;
	iq_etDiagExt	: PDL_ET_DiagExt;
	iq_sMsg			: STRING[80];
END_VAR

IF (iq_etDiag <> GD.ET_Diag.Ok) THEN
	CASE iq_etDiagExt OF

	PDL_ET_DiagExt.DriveInvalid: (* if Drive has no brake *)
		stExceptionModuleReaction2.etDiag := GD.ET_Diag.InputParameterInvalid;
		stExceptionModuleReaction2.udiDiagExt := AXM_ET_DiagExt.DriveInvalid;
		stExceptionModuleReaction2.sMsg := iq_sMsg;
		ReportException(iq_stException := stExceptionModuleReaction2);

	PDL_ET_DiagExt.DriveNotReady:
		stExceptionModuleReaction2.etDiag := GD.ET_Diag.DriveConditionInvalid;
		stExceptionModuleReaction2.udiDiagExt := AXM_ET_DiagExt.DriveNotReady;
		stExceptionModuleReaction2.sMsg := iq_sMsg;
		ReportException(iq_stException := stExceptionModuleReaction2);

	ELSE
		stExceptionUnexpected.udiDiagExt := AXM_ET_DiagExt.UnexpectedFeedback;
		stExceptionUnexpected.sMsg := SE_CTBX.FC_MultiConcat(	i_sString1 := 'FB_BrakeRelease ',
															i_sString2 := PDL_FC_EtDiagExtToString(i_etDiagExt := iq_etDiagExt),
															i_sString3 := ' ',
															i_sString4 := iq_sMsg);
		ReportException(iq_stException := stExceptionUnexpected);
	END_CASE
END_IF

(* ---- DiagTestDriveEnable.meth.st ---- *)
{attribute 'conditionalshow_all_locals'}
METHOD INTERNAL DiagTestDriveEnable
VAR_IN_OUT
	iq_etDiag		: GD.ET_Diag;
	iq_etDiagExt	: PDL_ET_DiagExt;
	iq_sMsg			: STRING[80];
END_VAR

IF (iq_etDiag <> GD.ET_Diag.Ok) THEN
	CASE iq_etDiagExt OF
	PDL_ET_DiagExt.DriveNotReady:
		stExceptionModuleReaction2.etDiag := GD.ET_Diag.DriveConditionInvalid;
		stExceptionModuleReaction2.udiDiagExt := AXM_ET_DiagExt.DriveNotReady;
		stExceptionModuleReaction2.sMsg := iq_sMsg;
		ReportException(iq_stException := stExceptionModuleReaction2);

	PDL_ET_DiagExt.InverterEnableOff:
		stExceptionModuleReaction2.etDiag := GD.ET_Diag.DriveConditionInvalid;
		stExceptionModuleReaction2.udiDiagExt := AXM_ET_DiagExt.InverterEnableOff;
		stExceptionModuleReaction2.sMsg := iq_sMsg;
		ReportException(iq_stException := stExceptionModuleReaction2);

	PDL_ET_DiagExt.TorqueEnableOff:
		stExceptionModuleReaction2.etDiag := GD.ET_Diag.DriveConditionInvalid;
		stExceptionModuleReaction2.udiDiagExt := AXM_ET_DiagExt.TorqueEnableOff;
		stExceptionModuleReaction2.sMsg := iq_sMsg;
		ReportException(iq_stException := stExceptionModuleReaction2);

	PDL_ET_DiagExt.PowerSupplyInvalid:
		stExceptionModuleReaction2.etDiag := GD.ET_Diag.InputParameterInvalid;
		stExceptionModuleReaction2.udiDiagExt := AXM_ET_DiagExt.PowerSupplyInvalid;
		stExceptionModuleReaction2.sMsg := iq_sMsg;
		ReportException(iq_stException := stExceptionModuleReaction2);

	PDL_ET_DiagExt.PowerSupplyNotFound:
		stExceptionModuleReaction2.etDiag := GD.ET_Diag.InputParameterInvalid;
		stExceptionModuleReaction2.udiDiagExt := AXM_ET_DiagExt.PowerSupplyNotFound;
		stExceptionModuleReaction2.sMsg := iq_sMsg;
		ReportException(iq_stException := stExceptionModuleReaction2);

	PDL_ET_DiagExt.PowerSupplyNotReady:
		stExceptionModuleReaction2.etDiag := GD.ET_Diag.PowerSupplyConditionInvalid;
		stExceptionModuleReaction2.udiDiagExt := AXM_ET_DiagExt.PowerSupplyNotReady;
		stExceptionModuleReaction2.sMsg := iq_sMsg;
		ReportException(iq_stException := stExceptionModuleReaction2);

	ELSE
		stExceptionUnexpected.udiDiagExt := AXM_ET_DiagExt.UnexpectedFeedback;
		stExceptionUnexpected.sMsg := SE_CTBX.FC_MultiConcat(	i_sString1 := 'FB_DriveEnable ',
															i_sString2 := PDL_FC_EtDiagExtToString(i_etDiagExt := iq_etDiagExt),
															i_sString3 := ' ',
															i_sString4 := iq_sMsg);
		ReportException(iq_stException := stExceptionUnexpected);
	END_CASE
END_IF

(* ---- DiagTestEndless.meth.st ---- *)
{attribute 'conditionalshow_all_locals'}
METHOD INTERNAL DiagTestEndless
VAR_IN_OUT
	iq_etDiag		: GD.ET_Diag;
	iq_etDiagExt	: PDL_ET_DiagExt;
	iq_sMsg			: STRING[80];
END_VAR

IF (iq_etDiag <> GD.ET_Diag.Ok) THEN
	CASE iq_etDiagExt OF
	PDL_ET_DiagExt.VelRange:
		stExceptionModuleReaction2.etDiag := GD.ET_Diag.InputParameterInvalid;
		stExceptionModuleReaction2.udiDiagExt := AXM_ET_DiagExt.VelRange;
		stExceptionModuleReaction2.sMsg := iq_sMsg;
		ReportException(iq_stException := stExceptionModuleReaction2);

	PDL_ET_DiagExt.AccRange:
		stExceptionModuleReaction2.etDiag := GD.ET_Diag.InputParameterInvalid;
		stExceptionModuleReaction2.udiDiagExt := AXM_ET_DiagExt.AccRange;
		stExceptionModuleReaction2.sMsg := iq_sMsg;
		ReportException(iq_stException := stExceptionModuleReaction2);

	PDL_ET_DiagExt.DecRange:
		stExceptionModuleReaction2.etDiag := GD.ET_Diag.InputParameterInvalid;
		stExceptionModuleReaction2.udiDiagExt := AXM_ET_DiagExt.DecRange;
		stExceptionModuleReaction2.sMsg := iq_sMsg;
		ReportException(iq_stException := stExceptionModuleReaction2);

	PDL_ET_DiagExt.JerkRange:
		stExceptionModuleReaction2.etDiag := GD.ET_Diag.InputParameterInvalid;
		stExceptionModuleReaction2.udiDiagExt := AXM_ET_DiagExt.JerkRange;
		stExceptionModuleReaction2.sMsg := iq_sMsg;
		ReportException(iq_stException := stExceptionModuleReaction2);

	PDL_ET_DiagExt.PeriodRange:
		stExceptionModuleReaction2.etDiag := GD.ET_Diag.InputParameterInvalid;
		stExceptionModuleReaction2.udiDiagExt := AXM_ET_DiagExt.PeriodRange;
		stExceptionModuleReaction2.sMsg := iq_sMsg;
		ReportException(iq_stException := stExceptionModuleReaction2);

	PDL_ET_DiagExt.StopPositionRange:
		stExceptionModuleReaction2.etDiag := GD.ET_Diag.InputParameterInvalid;
		stExceptionModuleReaction2.udiDiagExt := AXM_ET_DiagExt.StopPositionRange;
		stExceptionModuleReaction2.sMsg := iq_sMsg;
		ReportException(iq_stException := stExceptionModuleReaction2);

	ELSE
		stExceptionUnexpected.udiDiagExt := AXM_ET_DiagExt.UnexpectedFeedback;
		stExceptionUnexpected.sMsg := SE_CTBX.FC_MultiConcat(	i_sString1 := 'FB_Endless ',
															i_sString2 := PDL_FC_EtDiagExtToString(i_etDiagExt := iq_etDiagExt),
															i_sString3 := ' ',
															i_sString4 := iq_sMsg);
		ReportException(iq_stException := stExceptionUnexpected);
	END_CASE
END_IF

(* ---- DiagTestHoming.meth.st ---- *)
{attribute 'conditionalshow_all_locals'}
METHOD INTERNAL DiagTestHoming
VAR_IN_OUT
	iq_etDiag		: GD.ET_Diag;
	iq_etDiagExt	: PDL_ET_DiagExt;
	iq_sMsg			: STRING[80];
END_VAR

IF (iq_etDiag <> GD.ET_Diag.Ok) THEN
	CASE iq_etDiagExt OF
	PDL_ET_DiagExt.AbsEncOffsetRange:
		stExceptionModuleReaction2.etDiag := GD.ET_Diag.InputParameterInvalid;
		stExceptionModuleReaction2.udiDiagExt := AXM_ET_DiagExt.AbsEncOffsetRange;
		stExceptionModuleReaction2.sMsg := iq_sMsg;
		ReportException(iq_stException := stExceptionModuleReaction2);

	PDL_ET_DiagExt.AccRange:
		stExceptionModuleReaction2.etDiag := GD.ET_Diag.InputParameterInvalid;
		stExceptionModuleReaction2.udiDiagExt := AXM_ET_DiagExt.AccRange;
		stExceptionModuleReaction2.sMsg := iq_sMsg;
		ReportException(iq_stException := stExceptionModuleReaction2);

	PDL_ET_DiagExt.CheckSumInvalid:
		stExceptionModuleReaction2.etDiag := GD.ET_Diag.InputParameterInvalid;
		stExceptionModuleReaction2.udiDiagExt := AXM_ET_DiagExt.CheckSumInvalid;
		stExceptionModuleReaction2.sMsg := iq_sMsg;
		ReportException(iq_stException := stExceptionModuleReaction2);

	PDL_ET_DiagExt.DataNVRamInvalid:
		stExceptionModuleReaction2.etDiag := GD.ET_Diag.InputParameterInvalid;
		stExceptionModuleReaction2.udiDiagExt := AXM_ET_DiagExt.DataNVRamInvalid;
		stExceptionModuleReaction2.sMsg := iq_sMsg;
		ReportException(iq_stException := stExceptionModuleReaction2);

	PDL_ET_DiagExt.DecRange:
		stExceptionModuleReaction2.etDiag := GD.ET_Diag.InputParameterInvalid;
		stExceptionModuleReaction2.udiDiagExt := AXM_ET_DiagExt.DecRange;
		stExceptionModuleReaction2.sMsg := iq_sMsg;
		ReportException(iq_stException := stExceptionModuleReaction2);

	PDL_ET_DiagExt.DriveEncoderInvalid:
		stExceptionModuleReaction2.etDiag := GD.ET_Diag.DriveConditionInvalid;
		stExceptionModuleReaction2.udiDiagExt := AXM_ET_DiagExt.DriveEncoderInvalid;
		stExceptionModuleReaction2.sMsg := iq_sMsg;
		ReportException(iq_stException := stExceptionModuleReaction2);

	PDL_ET_DiagExt.LencInvalid:
		stExceptionModuleReaction2.etDiag := GD.ET_Diag.InputParameterInvalid;
		stExceptionModuleReaction2.udiDiagExt := AXM_ET_DiagExt.LencInvalid;
		stExceptionModuleReaction2.sMsg := iq_sMsg;
		ReportException(iq_stException := stExceptionModuleReaction2);

	PDL_ET_DiagExt.DriveIsMoving:
		stExceptionModuleReaction2.etDiag := GD.ET_Diag.DriveConditionInvalid;
		stExceptionModuleReaction2.udiDiagExt := AXM_ET_DiagExt.DriveIsMoving;
		stExceptionModuleReaction2.sMsg := iq_sMsg;
		ReportException(iq_stException := stExceptionModuleReaction2);

	PDL_ET_DiagExt.DriveNotDisabled:
		stExceptionModuleReaction2.etDiag := GD.ET_Diag.DriveConditionInvalid;
		stExceptionModuleReaction2.udiDiagExt := AXM_ET_DiagExt.DriveNotDisabled;
		stExceptionModuleReaction2.sMsg := iq_sMsg;
		ReportException(iq_stException := stExceptionModuleReaction2);

	PDL_ET_DiagExt.DriveNotReady:
		stExceptionModuleReaction2.etDiag := GD.ET_Diag.DriveConditionInvalid;
		stExceptionModuleReaction2.udiDiagExt := AXM_ET_DiagExt.DriveNotReady;
		stExceptionModuleReaction2.sMsg := iq_sMsg;
		ReportException(iq_stException := stExceptionModuleReaction2);

	PDL_ET_DiagExt.HwLimitNegReached:
		stExceptionModuleReaction2.etDiag := GD.ET_Diag.LimitReached;
		stExceptionModuleReaction2.udiDiagExt := AXM_ET_DiagExt.HwLimitNegReached;
		stExceptionModuleReaction2.sMsg := iq_sMsg;
		ReportException(iq_stException := stExceptionModuleReaction2);

	PDL_ET_DiagExt.HwLimitPosReached:
		stExceptionModuleReaction2.etDiag := GD.ET_Diag.LimitReached;
		stExceptionModuleReaction2.udiDiagExt := AXM_ET_DiagExt.HwLimitPosReached;
		stExceptionModuleReaction2.sMsg := iq_sMsg;
		ReportException(iq_stException := stExceptionModuleReaction2);

	PDL_ET_DiagExt.JerkRange:
		stExceptionModuleReaction2.etDiag := GD.ET_Diag.InputParameterInvalid;
		stExceptionModuleReaction2.udiDiagExt := AXM_ET_DiagExt.JerkRange;
		stExceptionModuleReaction2.sMsg := iq_sMsg;
		ReportException(iq_stException := stExceptionModuleReaction2);

	PDL_ET_DiagExt.LowVelRange:
		stExceptionModuleReaction2.etDiag := GD.ET_Diag.InputParameterInvalid;
		stExceptionModuleReaction2.udiDiagExt := AXM_ET_DiagExt.LowVelRange;
		stExceptionModuleReaction2.sMsg := iq_sMsg;
		ReportException(iq_stException := stExceptionModuleReaction2);

	PDL_ET_DiagExt.MaxTorqueNotFound:
		stExceptionModuleReaction2.etDiag := GD.ET_Diag.HomingFailed;
		stExceptionModuleReaction2.udiDiagExt := AXM_ET_DiagExt.MaxTorqueNotFound;
		stExceptionModuleReaction2.sMsg := iq_sMsg;
		ReportException(iq_stException := stExceptionModuleReaction2);

	PDL_ET_DiagExt.MaxTorqueRange:
		stExceptionModuleReaction2.etDiag := GD.ET_Diag.InputParameterInvalid;
		stExceptionModuleReaction2.udiDiagExt := AXM_ET_DiagExt.MaxTorqueRange;
		stExceptionModuleReaction2.sMsg := iq_sMsg;
		ReportException(iq_stException := stExceptionModuleReaction2);

	PDL_ET_DiagExt.MaxForceNotFound:
		stExceptionModuleReaction2.etDiag := GD.ET_Diag.HomingFailed;
		stExceptionModuleReaction2.udiDiagExt := AXM_ET_DiagExt.MaxForceNotFound;
		stExceptionModuleReaction2.sMsg := iq_sMsg;
		ReportException(iq_stException := stExceptionModuleReaction2);

	PDL_ET_DiagExt.MaxForceRange:
		stExceptionModuleReaction2.etDiag := GD.ET_Diag.InputParameterInvalid;
		stExceptionModuleReaction2.udiDiagExt := AXM_ET_DiagExt.MaxForceRange;
		stExceptionModuleReaction2.sMsg := iq_sMsg;
		ReportException(iq_stException := stExceptionModuleReaction2);

	PDL_ET_DiagExt.MaxTravelRange:
		stExceptionModuleReaction2.etDiag := GD.ET_Diag.InputParameterInvalid;
		stExceptionModuleReaction2.udiDiagExt := AXM_ET_DiagExt.MaxTravelRange;
		stExceptionModuleReaction2.sMsg := iq_sMsg;
		ReportException(iq_stException := stExceptionModuleReaction2);

	PDL_ET_DiagExt.NoAccessToEEPROM:
		stExceptionModuleReaction2.etDiag := GD.ET_Diag.DriveConditionInvalid;
		stExceptionModuleReaction2.udiDiagExt := AXM_ET_DiagExt.NoAccessToEEPROM;
		stExceptionModuleReaction2.sMsg := iq_sMsg;
		ReportException(iq_stException := stExceptionModuleReaction2);

	PDL_ET_DiagExt.PointerRestorePosRetainInvalid:
		stExceptionModuleReaction2.etDiag := GD.ET_Diag.InputParameterInvalid;
		stExceptionModuleReaction2.udiDiagExt := AXM_ET_DiagExt.PointerRestorePosRetainInvalid;
		stExceptionModuleReaction2.sMsg := iq_sMsg;
		ReportException(iq_stException := stExceptionModuleReaction2);

	PDL_ET_DiagExt.ProgrammingInProgress:
		stExceptionModuleReaction2.etDiag := GD.ET_Diag.DriveConditionInvalid;
		stExceptionModuleReaction2.udiDiagExt := AXM_ET_DiagExt.ProgrammingInProgress;
		stExceptionModuleReaction2.sMsg := iq_sMsg;
		ReportException(iq_stException := stExceptionModuleReaction2);

	PDL_ET_DiagExt.ProgrammingInvalidEEPROM:
		stExceptionModuleReaction2.etDiag := GD.ET_Diag.DriveConditionInvalid;
		stExceptionModuleReaction2.udiDiagExt := AXM_ET_DiagExt.ProgrammingInvalidEEPROM;
		stExceptionModuleReaction2.sMsg := iq_sMsg;
		ReportException(iq_stException := stExceptionModuleReaction2);

	PDL_ET_DiagExt.RestoreInterrupted:
		stExceptionModuleReaction2.etDiag := GD.ET_Diag.DriveConditionInvalid;
		stExceptionModuleReaction2.udiDiagExt := AXM_ET_DiagExt.RestoreInterrupted;
		stExceptionModuleReaction2.sMsg := iq_sMsg;
		ReportException(iq_stException := stExceptionModuleReaction2);

	PDL_ET_DiagExt.SensorNotFound:
		stExceptionModuleReaction2.etDiag := GD.ET_Diag.HomingFailed;
		stExceptionModuleReaction2.udiDiagExt := AXM_ET_DiagExt.SensorNotFound;
		stExceptionModuleReaction2.sMsg := iq_sMsg;
		ReportException(iq_stException := stExceptionModuleReaction2);

	PDL_ET_DiagExt.SercosNotInPhaseFour:
		stExceptionModuleReaction2.etDiag := GD.ET_Diag.SercosConditionInvalid;
		stExceptionModuleReaction2.udiDiagExt := AXM_ET_DiagExt.SercosNotInPhaseFour;
		stExceptionModuleReaction2.sMsg := iq_sMsg;
		ReportException(iq_stException := stExceptionModuleReaction2);

	PDL_ET_DiagExt.TouchProbeInvalid:
		stExceptionModuleReaction2.etDiag := GD.ET_Diag.InputParameterInvalid;
		stExceptionModuleReaction2.udiDiagExt := AXM_ET_DiagExt.TouchProbeInvalid;
		stExceptionModuleReaction2.sMsg := iq_sMsg;
		ReportException(iq_stException := stExceptionModuleReaction2);

	PDL_ET_DiagExt.TouchProbeNotActive:
		stExceptionModuleReaction2.etDiag := GD.ET_Diag.InputParameterInvalid;
		stExceptionModuleReaction2.udiDiagExt := AXM_ET_DiagExt.TouchProbeNotActive;
		stExceptionModuleReaction2.sMsg := iq_sMsg;
		ReportException(iq_stException := stExceptionModuleReaction2);

	PDL_ET_DiagExt.TouchProbeNotFound:
		stExceptionModuleReaction2.etDiag := GD.ET_Diag.HomingFailed;
		stExceptionModuleReaction2.udiDiagExt := AXM_ET_DiagExt.TouchProbeNotFound;
		stExceptionModuleReaction2.sMsg := iq_sMsg;
		ReportException(iq_stException := stExceptionModuleReaction2);

	PDL_ET_DiagExt.TouchProbeVirtual:
		stExceptionModuleReaction2.etDiag := GD.ET_Diag.InputParameterInvalid;
		stExceptionModuleReaction2.udiDiagExt := AXM_ET_DiagExt.TouchProbeVirtual;
		stExceptionModuleReaction2.sMsg := iq_sMsg;
		ReportException(iq_stException := stExceptionModuleReaction2);

	PDL_ET_DiagExt.UserPeriodRange:
		stExceptionModuleReaction2.etDiag := GD.ET_Diag.InputParameterInvalid;
		stExceptionModuleReaction2.udiDiagExt := AXM_ET_DiagExt.UserPeriodRange;
		stExceptionModuleReaction2.sMsg := iq_sMsg;
		ReportException(iq_stException := stExceptionModuleReaction2);

	PDL_ET_DiagExt.VelRange:
		stExceptionModuleReaction2.etDiag := GD.ET_Diag.InputParameterInvalid;
		stExceptionModuleReaction2.udiDiagExt := AXM_ET_DiagExt.VelRange;
		stExceptionModuleReaction2.sMsg := iq_sMsg;
		ReportException(iq_stException := stExceptionModuleReaction2);

	PDL_ET_DiagExt.UnknownMode:
		stExceptionModuleReaction2.etDiag := GD.ET_Diag.InputParameterInvalid;
		stExceptionModuleReaction2.udiDiagExt := AXM_ET_DiagExt.UnknownMode;
		stExceptionModuleReaction2.sMsg := iq_sMsg;
		ReportException(iq_stException := stExceptionModuleReaction2);

	PDL_ET_DiagExt.HwLimitNegStillActive:
		stExceptionModuleReaction2.etDiag := GD.ET_Diag.ExecutionAborted;
		stExceptionModuleReaction2.udiDiagExt := AXM_ET_DiagExt.HwLimitNegStillActive;
		stExceptionModuleReaction2.sMsg := iq_sMsg;
		ReportException(iq_stException := stExceptionModuleReaction2);

	PDL_ET_DiagExt.HwLimitPosStillActive:
		stExceptionModuleReaction2.etDiag := GD.ET_Diag.ExecutionAborted;
		stExceptionModuleReaction2.udiDiagExt := AXM_ET_DiagExt.HwLimitPosStillActive;
		stExceptionModuleReaction2.sMsg := iq_sMsg;
		ReportException(iq_stException := stExceptionModuleReaction2);

	PDL_ET_DiagExt.ReducedVelocityLImit:
		stExceptionModuleReaction2.etDiag := GD.ET_Diag.LimitReached;
		stExceptionModuleReaction2.udiDiagExt := AXM_ET_DiagExt.ReducedVelocityLImit;
		stExceptionModuleReaction2.sMsg := iq_sMsg;
		ReportException(iq_stException := stExceptionModuleReaction2);

	PDL_ET_DiagExt.ReducedVelocityRange:
		stExceptionModuleReaction2.etDiag := GD.ET_Diag.InputParameterInvalid;
		stExceptionModuleReaction2.udiDiagExt := AXM_ET_DiagExt.ReducedVelocityRange;
		stExceptionModuleReaction2.sMsg := iq_sMsg;
		ReportException(iq_stException := stExceptionModuleReaction2);

	PDL_ET_DiagExt.ReducedVelocityFactorRange:
		stExceptionModuleReaction2.etDiag := GD.ET_Diag.InputParameterInvalid;
		stExceptionModuleReaction2.udiDiagExt := AXM_ET_DiagExt.ReducedVelocityFactorRange;
		stExceptionModuleReaction2.sMsg := iq_sMsg;
		ReportException(iq_stException := stExceptionModuleReaction2);

	PDL_ET_DiagExt.OutOfRestoreWindow:
		stExceptionModuleReaction2.etDiag := GD.ET_Diag.LimitReached;
		stExceptionModuleReaction2.udiDiagExt := AXM_ET_DiagExt.OutOfRestoreWindow;
		stExceptionModuleReaction2.sMsg := iq_sMsg;
		ReportException(iq_stException := stExceptionModuleReaction2);

	ELSE
		stExceptionUnexpected.udiDiagExt := AXM_ET_DiagExt.UnexpectedFeedback;
		stExceptionUnexpected.sMsg := SE_CTBX.FC_MultiConcat(	i_sString1 := 'FB_Home ',
															i_sString2 := PDL_FC_EtDiagExtToString(i_etDiagExt := iq_etDiagExt),
															i_sString3 := ' ',
															i_sString4 := iq_sMsg);
		ReportException(iq_stException := stExceptionUnexpected);
	END_CASE
END_IF

(* ---- DiagTestJogging.meth.st ---- *)
{attribute 'conditionalshow_all_locals'}
METHOD INTERNAL DiagTestJogging
VAR_IN_OUT
	iq_etDiag		: GD.ET_Diag;
	iq_etDiagExt	: PDL_ET_DiagExt;
	iq_sMsg			: STRING[80];
END_VAR

IF (iq_etDiag <> GD.ET_Diag.Ok) THEN
	CASE iq_etDiagExt OF
	PDL_ET_DiagExt.VelRange:
		stExceptionModuleReaction2.etDiag := GD.ET_Diag.InputParameterInvalid;
		stExceptionModuleReaction2.udiDiagExt := AXM_ET_DiagExt.VelRange;
		stExceptionModuleReaction2.sMsg := iq_sMsg;
		ReportException(iq_stException := stExceptionModuleReaction2);

	PDL_ET_DiagExt.AccRange:
		stExceptionModuleReaction2.etDiag := GD.ET_Diag.InputParameterInvalid;
		stExceptionModuleReaction2.udiDiagExt := AXM_ET_DiagExt.AccRange;
		stExceptionModuleReaction2.sMsg := iq_sMsg;
		ReportException(iq_stException := stExceptionModuleReaction2);

	PDL_ET_DiagExt.DecRange:
		stExceptionModuleReaction2.etDiag := GD.ET_Diag.InputParameterInvalid;
		stExceptionModuleReaction2.udiDiagExt := AXM_ET_DiagExt.DecRange;
		stExceptionModuleReaction2.sMsg := iq_sMsg;
		ReportException(iq_stException := stExceptionModuleReaction2);

	PDL_ET_DiagExt.JerkRange:
		stExceptionModuleReaction2.etDiag := GD.ET_Diag.InputParameterInvalid;
		stExceptionModuleReaction2.udiDiagExt := AXM_ET_DiagExt.JerkRange;
		stExceptionModuleReaction2.sMsg := iq_sMsg;
		ReportException(iq_stException := stExceptionModuleReaction2);

	PDL_ET_DiagExt.MaxDistanceRange:
		stExceptionModuleReaction2.etDiag := GD.ET_Diag.InputParameterInvalid;
		stExceptionModuleReaction2.udiDiagExt := AXM_ET_DiagExt.MaxDistanceRange;
		stExceptionModuleReaction2.sMsg := iq_sMsg;
		ReportException(iq_stException := stExceptionModuleReaction2);

	PDL_ET_DiagExt.PeriodRange:
		stExceptionModuleReaction2.etDiag := GD.ET_Diag.InputParameterInvalid;
		stExceptionModuleReaction2.udiDiagExt := AXM_ET_DiagExt.PeriodRange;
		stExceptionModuleReaction2.sMsg := iq_sMsg;
		ReportException(iq_stException := stExceptionModuleReaction2);

	ELSE
		stExceptionUnexpected.udiDiagExt := AXM_ET_DiagExt.UnexpectedFeedback;
		stExceptionUnexpected.sMsg := SE_CTBX.FC_MultiConcat(	i_sString1 := 'FB_Jogging ',
															i_sString2 := PDL_FC_EtDiagExtToString(i_etDiagExt := iq_etDiagExt),
															i_sString3 := ' ',
															i_sString4 := iq_sMsg);
		ReportException(iq_stException := stExceptionUnexpected);
	END_CASE
END_IF

(* ---- DiagTestMultiCam.meth.st ---- *)
{attribute 'conditionalshow_all_locals'}
METHOD INTERNAL DiagTestMultiCam
VAR_IN_OUT
	iq_etDiag		: GD.ET_Diag;
	iq_etDiagExt	: PDL_ET_DiagExt;
	iq_sMsg			: STRING[80];
END_VAR

IF (iq_etDiag <> GD.ET_Diag.Ok) THEN
	CASE iq_etDiagExt OF
	PDL_ET_DiagExt.AccRange:
		stExceptionModuleReaction2.etDiag := GD.ET_Diag.InputParameterInvalid;
		stExceptionModuleReaction2.udiDiagExt := AXM_ET_DiagExt.AccRange;
		stExceptionModuleReaction2.sMsg := iq_sMsg;
		ReportException(iq_stException := stExceptionModuleReaction2);

	PDL_ET_DiagExt.BoundaryConditionInvalid:
		stExceptionModuleReaction2.etDiag := GD.ET_Diag.InputParameterInvalid;
		stExceptionModuleReaction2.udiDiagExt := AXM_ET_DiagExt.BoundaryConditionInvalid;
		stExceptionModuleReaction2.sMsg := iq_sMsg;
		ReportException(iq_stException := stExceptionModuleReaction2);

	PDL_ET_DiagExt.DecRange:
		stExceptionModuleReaction2.etDiag := GD.ET_Diag.InputParameterInvalid;
		stExceptionModuleReaction2.udiDiagExt := AXM_ET_DiagExt.DecRange;
		stExceptionModuleReaction2.sMsg := iq_sMsg;
		ReportException(iq_stException := stExceptionModuleReaction2);

	PDL_ET_DiagExt.JerkRange:
		stExceptionModuleReaction2.etDiag := GD.ET_Diag.InputParameterInvalid;
		stExceptionModuleReaction2.udiDiagExt := AXM_ET_DiagExt.JerkRange;
		stExceptionModuleReaction2.sMsg := iq_sMsg;
		ReportException(iq_stException := stExceptionModuleReaction2);

	PDL_ET_DiagExt.NumberOfCamPointsRange:
		stExceptionModuleReaction2.etDiag := GD.ET_Diag.InputParameterInvalid;
		stExceptionModuleReaction2.udiDiagExt := AXM_ET_DiagExt.NumberOfCamPointsRange;
		stExceptionModuleReaction2.sMsg := iq_sMsg;
		ReportException(iq_stException := stExceptionModuleReaction2);

	PDL_ET_DiagExt.RangeK:
		stExceptionModuleReaction2.etDiag := GD.ET_Diag.InputParameterInvalid;
		stExceptionModuleReaction2.udiDiagExt := AXM_ET_DiagExt.RangeK;
		stExceptionModuleReaction2.sMsg := iq_sMsg;
		ReportException(iq_stException := stExceptionModuleReaction2);

	PDL_ET_DiagExt.RangeM:
		stExceptionModuleReaction2.etDiag := GD.ET_Diag.InputParameterInvalid;
		stExceptionModuleReaction2.udiDiagExt := AXM_ET_DiagExt.RangeM;
		stExceptionModuleReaction2.sMsg := iq_sMsg;
		ReportException(iq_stException := stExceptionModuleReaction2);

	PDL_ET_DiagExt.UnknownCamType:
		stExceptionModuleReaction2.etDiag := GD.ET_Diag.InputParameterInvalid;
		stExceptionModuleReaction2.udiDiagExt := AXM_ET_DiagExt.UnknownCamType;
		stExceptionModuleReaction2.sMsg := iq_sMsg;
		ReportException(iq_stException := stExceptionModuleReaction2);

	PDL_ET_DiagExt.UnknownCsModeMaster:
		stExceptionModuleReaction2.etDiag := GD.ET_Diag.InputParameterInvalid;
		stExceptionModuleReaction2.udiDiagExt := AXM_ET_DiagExt.UnknownCsModeMaster;
		stExceptionModuleReaction2.sMsg := iq_sMsg;
		ReportException(iq_stException := stExceptionModuleReaction2);

	PDL_ET_DiagExt.UnknownCsModeSlave:
		stExceptionModuleReaction2.etDiag := GD.ET_Diag.InputParameterInvalid;
		stExceptionModuleReaction2.udiDiagExt := AXM_ET_DiagExt.UnknownCsModeSlave;
		stExceptionModuleReaction2.sMsg := iq_sMsg;
		ReportException(iq_stException := stExceptionModuleReaction2);

	PDL_ET_DiagExt.UnknownWsMode:
		stExceptionModuleReaction2.etDiag := GD.ET_Diag.InputParameterInvalid;
		stExceptionModuleReaction2.udiDiagExt := AXM_ET_DiagExt.UnknownWsMode;
		stExceptionModuleReaction2.sMsg := iq_sMsg;
		ReportException(iq_stException := stExceptionModuleReaction2);

	PDL_ET_DiagExt.VelRange:
		stExceptionModuleReaction2.etDiag := GD.ET_Diag.InputParameterInvalid;
		stExceptionModuleReaction2.udiDiagExt := AXM_ET_DiagExt.VelRange;
		stExceptionModuleReaction2.sMsg := iq_sMsg;
		ReportException(iq_stException := stExceptionModuleReaction2);

	PDL_ET_DiagExt.XFactorTooSmall:
		stExceptionModuleReaction2.etDiag := GD.ET_Diag.InputParameterInvalid;
		stExceptionModuleReaction2.udiDiagExt := AXM_ET_DiagExt.XFactorTooLow;
		stExceptionModuleReaction2.sMsg := iq_sMsg;
		ReportException(iq_stException := stExceptionModuleReaction2);

	PDL_ET_DiagExt.YEqualCheckFailed:
		stExceptionModuleReaction2.etDiag := GD.ET_Diag.InputParameterInvalid;
		stExceptionModuleReaction2.udiDiagExt := AXM_ET_DiagExt.YEqualCheckFailed;
		stExceptionModuleReaction2.sMsg := iq_sMsg;
		ReportException(iq_stException := stExceptionModuleReaction2);

	PDL_ET_DiagExt.DrivePositionOutOfWsWindow:
		stExceptionModuleReaction2.etDiag := GD.ET_Diag.WarmStartConditionInvalid;
		stExceptionModuleReaction2.udiDiagExt := AXM_ET_DiagExt.DrivePositionOutOfWsWindow;
		stExceptionModuleReaction2.sMsg := iq_sMsg;
		ReportException(iq_stException := stExceptionModuleReaction2);

	PDL_ET_DiagExt.MasterMoved:
		stExceptionModuleReaction2.etDiag := GD.ET_Diag.WarmStartConditionInvalid;
		stExceptionModuleReaction2.udiDiagExt := AXM_ET_DiagExt.MasterMoved;
		stExceptionModuleReaction2.sMsg := iq_sMsg;
		ReportException(iq_stException := stExceptionModuleReaction2);

	PDL_ET_DiagExt.UserCamHasBeenDeleted:
		stExceptionModuleReaction2.etDiag := GD.ET_Diag.WarmStartConditionInvalid;
		stExceptionModuleReaction2.udiDiagExt := AXM_ET_DiagExt.UserCamHasBeenDeleted;
		stExceptionModuleReaction2.sMsg := iq_sMsg;
		ReportException(iq_stException := stExceptionModuleReaction2);

	ELSE
		stExceptionUnexpected.udiDiagExt := AXM_ET_DiagExt.UnexpectedFeedback;
		stExceptionUnexpected.sMsg := SE_CTBX.FC_MultiConcat(	i_sString1 := 'FB_MultiCam ',
															i_sString2 := PDL_FC_EtDiagExtToString(i_etDiagExt := iq_etDiagExt),
															i_sString3 := ' ',
															i_sString4 := iq_sMsg);
		ReportException(iq_stException := stExceptionUnexpected);
	END_CASE
END_IF

(* ---- DiagTestPositioning.meth.st ---- *)
{attribute 'conditionalshow_all_locals'}
METHOD INTERNAL DiagTestPositioning
VAR_IN_OUT
	iq_etDiag		: GD.ET_Diag;
	iq_etDiagExt	: PDL_ET_DiagExt;
	iq_sMsg			: STRING[80];
END_VAR

IF (iq_etDiag <> GD.ET_Diag.Ok) THEN
	CASE iq_etDiagExt OF
	PDL_ET_DiagExt.AccRange:
		stExceptionModuleReaction2.etDiag := GD.ET_Diag.InputParameterInvalid;
		stExceptionModuleReaction2.udiDiagExt := AXM_ET_DiagExt.AccRange;
		stExceptionModuleReaction2.sMsg := iq_sMsg;
		ReportException(iq_stException := stExceptionModuleReaction2);

	PDL_ET_DiagExt.DecRange:
		stExceptionModuleReaction2.etDiag := GD.ET_Diag.InputParameterInvalid;
		stExceptionModuleReaction2.udiDiagExt := AXM_ET_DiagExt.DecRange;
		stExceptionModuleReaction2.sMsg := iq_sMsg;
		ReportException(iq_stException := stExceptionModuleReaction2);

	PDL_ET_DiagExt.JerkRange:
		stExceptionModuleReaction2.etDiag := GD.ET_Diag.InputParameterInvalid;
		stExceptionModuleReaction2.udiDiagExt := AXM_ET_DiagExt.JerkRange;
		stExceptionModuleReaction2.sMsg := iq_sMsg;
		ReportException(iq_stException := stExceptionModuleReaction2);

	PDL_ET_DiagExt.VelRange:
		stExceptionModuleReaction2.etDiag := GD.ET_Diag.InputParameterInvalid;
		stExceptionModuleReaction2.udiDiagExt := AXM_ET_DiagExt.VelRange;
		stExceptionModuleReaction2.sMsg := iq_sMsg;
		ReportException(iq_stException := stExceptionModuleReaction2);

	PDL_ET_DiagExt.PosModeRange:
		stExceptionModuleReaction2.etDiag := GD.ET_Diag.InputParameterInvalid;
		stExceptionModuleReaction2.udiDiagExt := AXM_ET_DiagExt.PosModeRange;
		stExceptionModuleReaction2.sMsg := iq_sMsg;
		ReportException(iq_stException := stExceptionModuleReaction2);

	ELSE
		stExceptionUnexpected.udiDiagExt := AXM_ET_DiagExt.UnexpectedFeedback;
		stExceptionUnexpected.sMsg := SE_CTBX.FC_MultiConcat(	i_sString1 := 'fbPos ',
															i_sString2 := PDL_FC_EtDiagExtToString(i_etDiagExt := iq_etDiagExt),
															i_sString3 := ' ',
															i_sString4 := iq_sMsg);
		ReportException(iq_stException := stExceptionUnexpected);
	END_CASE
END_IF

(* ---- DisableAllJobs.meth.st ---- *)
{attribute 'conditionalshow_all_locals'}
METHOD INTERNAL DisableAllJobs
VAR_INPUT
END_VAR

(* OpModes *)
	xRefEnable := FALSE;
	xManEnable := FALSE;
	xCamEnable := FALSE;
	xEndlessEnable := FALSE;
	xPosEnable := FALSE;
	xBrakeEnable := FALSE;
	xAdditionalEnable := FALSE;

(* ---- Endless_active.act.st ---- *)
__METADATA__
{
  "v3Meta": {
    "objectGuid": "3c0b60bf-17fe-403b-b7bd-421c8472aa89",
    "objectTypeGuid": "8ac092e5-3128-4e26-9e7e-11016c6684f2",
    "embeddedObjectTypeGuids": [
      "3b83b776-fb25-43b8-99f2-3c507c9143fc"
    ],
    "properties": {},
    "subObjects": {}
  }
}

iq_stAxisModuleItf.stMain.q_etOpMode := AXM_ET_OpMode.Endless;

IF (iq_stAxisModuleItf.stMain.stReducedVelocity.i_xEnableReducedVelocity AND
	NOT iq_stAxisModuleItf.stMain.stReducedVelocity.i_xOnlyLimitCheck) THEN

	lrEndlessVel := MIN(iq_stAxisModuleItf.stEndless.i_lrVel, iq_stAxisModuleItf.stMain.stReducedVelocity.i_lrMaxReducedVelocity);
ELSE
	lrEndlessVel := iq_stAxisModuleItf.stEndless.i_lrVel;
END_IF

xEndlessStart := (xStartFlag OR iq_stAxisModuleItf.stMain.i_xStart) AND NOT stModuleReaction.axReaction[TPL.ET_Reaction.StopEndOfCycle];

fbEndless(	i_xEnable			:= xEndlessEnable AND fbDriveEnable.q_xDriveEnabled,
			i_ifDrive			:= iq_stAxisModuleItf.stMain.i_ifDrive,
			i_lrVel				:= lrEndlessVel,
			i_lrAcc				:= iq_stAxisModuleItf.stEndless.i_lrAcc,
			i_lrDec				:= iq_stAxisModuleItf.stEndless.i_lrDec,
			i_lrJerk			:= iq_stAxisModuleItf.stEndless.i_lrJerk,
			i_lrPeriod			:= iq_stAxisModuleItf.stEndless.i_lrPeriod,
			i_lrStopPosition	:= iq_stAxisModuleItf.stEndless.i_lrStopPosition,
			i_xStart			:= xEndlessStart,
			q_etDiag			=> etDiagBuffer,
			q_etDiagExt			=> etDiagExtBufferPDL,
			q_sMsg				=> sDiagMsgBuffer,
			q_xInVelocity		=> iq_stAxisModuleItf.stEndless.q_xInVelocity);

DiagTestEndless(iq_etDiag		:= fbEndless.q_etDiag,
				iq_etDiagExt	:= fbEndless.q_etDiagExt,
				iq_sMsg			:= fbEndless.q_sMsg);

IF fbEndless.q_xReady AND fbEndless.q_etDiagExt = PDL_ET_DiagExt.WaitForStart THEN
	 iq_stAxisModuleItf.stMain.q_etState := AXM_ET_State.EndlessWaitForStart;
ELSIF fbEndless.q_xReady THEN
	iq_stAxisModuleItf.stMain.q_etState := AXM_ET_State.EndlessRunning;
ELSE
	IF xEndlessEnable THEN
		iq_stAxisModuleItf.stMain.q_etState := AXM_ET_State.EndlessInit;
	ELSE
		iq_stAxisModuleItf.stMain.q_etState := AXM_ET_State.EndlessExit;
	END_IF
END_IF

IF NOT xEndlessEnable AND NOT fbEndless.q_xActive THEN
	xEndlessActive := FALSE;
END_IF

(* ---- ExceptionHandler_active.act.st ---- *)
__METADATA__
{
  "v3Meta": {
    "objectGuid": "027a414b-2e1b-4ec2-826d-53250118d89b",
    "objectTypeGuid": "8ac092e5-3128-4e26-9e7e-11016c6684f2",
    "embeddedObjectTypeGuids": [
      "3b83b776-fb25-43b8-99f2-3c507c9143fc"
    ],
    "properties": {},
    "subObjects": {}
  }
}

IF iq_stStandardModuleItf.q_xActive THEN

(* -----------------------------------------------------------------------------------------------*)
(* Check Axis Exceptions *)
(* -----------------------------------------------------------------------------------------------*)
	GetInterfaces();
	IF ifDiagnostic <> 0 THEN
		IF (ifDiagnostic.DiagClass > 0)  AND (ifDiagnostic.DiagClass < 3) THEN
			sDiagMsgExt := ifDiagnostic.DiagExtMsg;
			stWarningDrive.sMsg := SE_CTBX.FC_MultiConcat(	i_sString1 := Standard.CONCAT('DiagCode: ', DINT_TO_STRING(ifDiagnostic.DiagCode)),
														i_sString2 := Standard.CONCAT(' Msg: ', ifDiagnostic.DiagMsg),
														i_sString3 := ' Ext: ',
														i_sString4 := sDiagMsgExt);
			stWarningDrive.udiExceptionNumber := TPL.FC_GenerateExceptionNumber(	i_etSource		:= TPL.ET_ExceptionSource.System,
																					i_udiDiagExt	:= DINT_TO_UDINT(ifDiagnostic.DiagCode),
																					q_etDiag		=> , // function has no errors
																					q_etDiagExt		=> );
			ReportException(iq_stException := stWarningDrive);
		END_IF
		IF (ifDiagnostic.DiagClass = 3) THEN
			sDiagMsgExt := ifDiagnostic.DiagExtMsg;
			stExcepitonDrive.sMsg := SE_CTBX.FC_MultiConcat(	i_sString1 := Standard.CONCAT('DiagCode: ', DINT_TO_STRING(ifDiagnostic.DiagCode)),
															i_sString2 := Standard.CONCAT(' Msg: ', ifDiagnostic.DiagMsg),
															i_sString3 := ' Ext: ',
															i_sString4 := sDiagMsgExt);
			stExcepitonDrive.udiExceptionNumber := TPL.FC_GenerateExceptionNumber(	i_etSource		:= TPL.ET_ExceptionSource.System,
																					i_udiDiagExt	:= DINT_TO_UDINT(ifDiagnostic.DiagCode),
																					q_etDiag		=> , // function has no errors
																					q_etDiagExt		=> );
			ReportException(iq_stException := stExcepitonDrive);
		END_IF
		IF (ifDiagnostic.DiagClass > 3) THEN
			sDiagMsgExt := ifDiagnostic.DiagExtMsg;
			stExceptionDriveFatal.sMsg := SE_CTBX.FC_MultiConcat(	i_sString1 := Standard.CONCAT('DiagCode: ', DINT_TO_STRING(ifDiagnostic.DiagCode)),
																i_sString2 := Standard.CONCAT(' Msg: ', ifDiagnostic.DiagMsg),
																i_sString3 := ' Ext: ',
																i_sString4 := sDiagMsgExt);
			stExceptionDriveFatal.udiExceptionNumber := TPL.FC_GenerateExceptionNumber(	i_etSource		:= TPL.ET_ExceptionSource.System,
																						i_udiDiagExt	:= DINT_TO_UDINT(ifDiagnostic.DiagCode),
																						q_etDiag		=> , // function has no errors
																						q_etDiagExt		=> );
			ReportException(iq_stException := stExceptionDriveFatal);
		END_IF
	ELSE
		sDiagMsgExt := '';
	END_IF

(* -----------------------------------------------------------------------------------------------*)
(* HW Limitswitches *)
(* -----------------------------------------------------------------------------------------------*)

	IF iq_stAxisModuleItf.stMain.i_xHwLimitPos AND
		(iq_stAxisModuleItf.stMain.q_etOpMode = AXM_ET_OpMode.MultiCam OR
		iq_stAxisModuleItf.stMain.q_etOpMode = AXM_ET_OpMode.Endless OR
		iq_stAxisModuleItf.stMain.q_etOpMode = AXM_ET_OpMode.Positioning OR
		iq_stAxisModuleItf.stMain.q_etOpMode = AXM_ET_OpMode.Additional) THEN

		ReportException(iq_stException := stExceptionPosHwLimit);

	ELSIF iq_stAxisModuleItf.stMain.i_xHwLimitPos AND
			iq_stAxisModuleItf.stMain.q_etOpMode = AXM_ET_OpMode.Homing AND
			(iq_stAxisModuleItf.stHome.i_etMode = PDL_ET_HomeMode.PosDirectionPosEdgeHWLimitPos OR
			 iq_stAxisModuleItf.stHome.i_etMode = PDL_ET_HomeMode.PosDirectionNegEdgeHWLimitPos) THEN
		; //do nothing and ignore HW-Limit Sensor
	ELSIF iq_stAxisModuleItf.stMain.i_xHwLimitPos AND (iq_stAxisModuleItf.stMain.q_etOpMode <> AXM_ET_OpMode.NoOp) THEN
		ReportException(iq_stException := stWarningPosHwLimit);
	ELSIF NOT iq_stAxisModuleItf.stMain.i_xHwLimitPos THEN
		CancelException(iq_stException := stWarningPosHwLimit);
	END_IF

	IF iq_stAxisModuleItf.stMain.i_xHwLimitNeg AND
		(iq_stAxisModuleItf.stMain.q_etOpMode = AXM_ET_OpMode.MultiCam OR
		iq_stAxisModuleItf.stMain.q_etOpMode = AXM_ET_OpMode.Endless OR
		iq_stAxisModuleItf.stMain.q_etOpMode = AXM_ET_OpMode.Positioning OR
		iq_stAxisModuleItf.stMain.q_etOpMode = AXM_ET_OpMode.Additional) THEN

		ReportException(iq_stException := stExceptionNegHwLimit);

	ELSIF iq_stAxisModuleItf.stMain.i_xHwLimitNeg AND
			iq_stAxisModuleItf.stMain.q_etOpMode = AXM_ET_OpMode.Homing AND
			(iq_stAxisModuleItf.stHome.i_etMode = PDL_ET_HomeMode.NegDirectionPosEdgeHWLimitNeg OR
			 iq_stAxisModuleItf.stHome.i_etMode = PDL_ET_HomeMode.NegDirectionNegEdgeHWLimitNeg) THEN
		; //do nothing and ignore HW-Limit Sensor
	ELSIF iq_stAxisModuleItf.stMain.i_xHwLimitNeg AND (iq_stAxisModuleItf.stMain.q_etOpMode <> AXM_ET_OpMode.NoOp) THEN
		ReportException(iq_stException := stWarningNegHwLimit);
	ELSIF NOT iq_stAxisModuleItf.stMain.i_xHwLimitNeg THEN
		CancelException(iq_stException := stWarningNegHwLimit);
	END_IF

(* -----------------------------------------------------------------------------------------------*)
(* Check Axis MechVelocity / ReducedVelocity *)
(* -----------------------------------------------------------------------------------------------*)
	IF iq_stAxisModuleItf.stMain.stReducedVelocity.i_xEnableReducedVelocity THEN

		IF ifDrive <> 0 THEN
			IF ABS(ifDrive.ActualPosition) > ABS(iq_stAxisModuleItf.stMain.stReducedVelocity.i_lrMaxReducedVelocity * iq_stAxisModuleItf.stMain.stReducedVelocity.i_lrReducedVelocityCheckFactor) THEN
					stExceptionVelLimitCrossed.sMsg := Standard.CONCAT('Vel: ', LREAL_TO_STRING(ifDrive.ActualVelocity));
					ReportException(iq_stException := stExceptionVelLimitCrossed);
			END_IF
		END_IF

	ELSE
		xInitReducedVel := FALSE;
	END_IF

(* -----------------------------------------------------------------------------------------------*)
(* Check StartPositionSelect (SCR#1459) *)
(* -----------------------------------------------------------------------------------------------*)
	IF iq_stAxisModuleItf.stMultiCam.iq_stExt.xStartPositionSelect THEN
		stExceptionModuleReaction2.etDiag := GD.ET_Diag.InputParameterInvalid;
		stExceptionModuleReaction2.udiDiagExt := AXM_ET_DiagExt.StartPositionSelectInvalid;
		stExceptionModuleReaction2.sMsg := 'xStartPositionSelect has to be false';
		ReportException(iq_stException := stExceptionModuleReaction2);
	END_IF

(* -----------------------------------------------------------------------------------------------*)
(* Check StopModi *)
(* -----------------------------------------------------------------------------------------------*)
(******* Reaction TPL.ET_Reaction.AsyncStop ********)
	IF stModuleReaction.axReaction[TPL.ET_Reaction.AsyncStop] THEN				(* Stop with ControllerStopt *)
		xCMDPowerOn := FALSE;
		IF NOT (xBrakeActive OR xBrakeEnable) THEN
			xStartFlag := FALSE;
			DisableAllJobs();
		END_IF
		xWsStartFlag := FALSE;

(******* Reaction TPL.ET_Reaction.SyncStopEL and TPL.ET_Reaction.SyncStopEH ********)
	ELSIF stModuleReaction.axReaction[TPL.ET_Reaction.SyncStopEH] OR stModuleReaction.axReaction[TPL.ET_Reaction.SyncStopEL] THEN
		fbTimeOut(IN:=TRUE, PT:= iq_stAxisModuleItf.stMain.i_timMasterStop);
		IF (iq_stAxisModuleItf.stMain.i_ifMaster <> 0) AND (iq_stAxisModuleItf.stMain.q_etOpMode = AXM_ET_OpMode.MultiCam) THEN
			lrMasterVel := GetMasterVel();
			IF (ABS(lrMasterVel) < 0.5 ) OR  fbTimeOut.Q THEN			(* Wait for Master stop or Timeout *)
				(* we have to wait until delay between master and slave caused by the deadtime is over,
					bevore we can disable the slaves cam job.
					Otherwise it would stop "asynchron" meaning, not completely synchron *)
				fbSyncStopDeadTimeDelay(IN:= TRUE, PT :=  T#2MS(*2ms = 2x sercos cycle time*));
				(* deadtime until the ref position (in the plc configuration) is up to date (= has taken the value it
				should have according to master.RefPosition*CAM) is 1 sercos cycle, to be on the secure side we wait
				2 sercos cylces, also because we don't test for refVelocity = 0 but < 0.5 *)
				IF(fbSyncStopDeadTimeDelay.Q OR fbTimeOut.Q) THEN
					(* synchron stop done and deadtime is over, or timeout (of IFB_TimeOut) *)
					IF NOT xBrakeActive AND NOT xBrakeEnable THEN
						xStartFlag := FALSE;
						xWsStartFlag := FALSE;
						DisableAllJobs();
					(* Reaction TPL.ET_Reaction.SyncStopEL *)
						IF stModuleReaction.axReaction[TPL.ET_Reaction.SyncStopEL] THEN
							xCMDPowerOn := FALSE;
						END_IF
					END_IF
				END_IF
			END_IF
		ELSE
		(*** immediately reaction if no master was found ***)
			IF NOT xBrakeActive AND NOT xBrakeEnable THEN
				xStartFlag := FALSE;
				xWsStartFlag := FALSE;
				DisableAllJobs();
				IF fbTimeOut.Q OR
					(iq_stAxisModuleItf.stMain.q_etOpMode = AXM_ET_OpMode.NoOp) THEN
					(* Reaction TPL.ET_Reaction.SyncStopEL *)
					IF stModuleReaction.axReaction[TPL.ET_Reaction.SyncStopEL] THEN
						xCMDPowerOn := FALSE;
					END_IF
				END_IF
			END_IF
		END_IF

(******* Reaction TPL.ET_Reaction.StopEndOfCycle ********)
	ELSIF stModuleReaction.axReaction[TPL.ET_Reaction.StopEndOfCycle] THEN
		IF NOT xCamActive AND NOT xBrakeActive THEN
			xStartFlag := FALSE;
			xWsStartFlag := FALSE;
		END_IF
	ELSE
		fbTimeOut(IN:= FALSE);
		fbSyncStopDeadTimeDelay(IN := FALSE);
	END_IF

END_IF

(* ---- GetInterfaces.act.st ---- *)
__METADATA__
{
  "v3Meta": {
    "objectGuid": "d17f2152-ffc0-400a-95a5-caef054ae84b",
    "objectTypeGuid": "8ac092e5-3128-4e26-9e7e-11016c6684f2",
    "embeddedObjectTypeGuids": [
      "3b83b776-fb25-43b8-99f2-3c507c9143fc"
    ],
    "properties": {},
    "subObjects": {}
  }
}

IF 	(iq_stAxisModuleItf.stMain.i_ifDrive <> 0) THEN
	IF (ifAxisOld <> iq_stAxisModuleItf.stMain.i_ifDrive) THEN
		ifAxisOld := iq_stAxisModuleItf.stMain.i_ifDrive;
		xSuccess := __QUERYINTERFACE(iq_stAxisModuleItf.stMain.i_ifDrive, ifGetParentDevice);
		IF xSuccess THEN
			ifDeviceAccess := ifGetParentDevice.GetParentDevice();
			xSuccess := __QUERYINTERFACE(ifDeviceAccess, ifDiagnosticAccess);
			IF xSuccess THEN
				ifDiagnostic := ifDiagnosticAccess.Diagnostic;
			END_IF
			xSuccess := __QUERYINTERFACE(ifDeviceAccess, ifDrive2Access);
			IF xSuccess THEN
				ifDrive2 := ifDrive2Access.Drive2;
			END_IF
			xSuccess := __QUERYINTERFACE(ifDeviceAccess, ifDriveAccess);
			IF xSuccess THEN
				ifDrive := ifDriveAccess.Drive;
			END_IF
		END_IF
	END_IF
END_IF

(* ---- GetMasterPosition.meth.st ---- *)
{attribute 'conditionalshow_all_locals'}
METHOD INTERNAL GetMasterPosition: LREAL
VAR_INPUT
END_VAR
VAR
END_VAR

GetMasterPosition := 0.0;

IF (iq_stAxisModuleItf.stMain.i_ifMaster <> 0) THEN
	GetMasterPosition := iq_stAxisModuleItf.stMain.i_ifMaster.lrPosition;
END_IF

(* ---- GetMasterVel.meth.st ---- *)
METHOD INTERNAL GetMasterVel : LREAL
VAR_INPUT
END_VAR
VAR

END_VAR

GetMasterVel := 0.0;

IF (iq_stAxisModuleItf.stMain.i_ifMaster <> 0) THEN
	GetMasterVel := iq_stAxisModuleItf.stMain.i_ifMaster.RefVelocity;
END_IF

(* ---- Homing_active.act.st ---- *)
__METADATA__
{
  "v3Meta": {
    "objectGuid": "efbee110-d1de-4db7-a717-9c786137436a",
    "objectTypeGuid": "8ac092e5-3128-4e26-9e7e-11016c6684f2",
    "embeddedObjectTypeGuids": [
      "3b83b776-fb25-43b8-99f2-3c507c9143fc"
    ],
    "properties": {},
    "subObjects": {}
  }
}

iq_stAxisModuleItf.stMain.q_etOpMode := AXM_ET_OpMode.Homing;
xRefStart := (xStartFlag OR iq_stAxisModuleItf.stMain.i_xStart) AND NOT stModuleReaction.axReaction[TPL.ET_Reaction.StopEndOfCycle];

fbHome.stReducedVelocity := iq_stAxisModuleItf.stMain.stReducedVelocity;
CASE iq_stAxisModuleItf.stHome.i_etMode OF
	PDL_ET_HomeMode.PosDirectionPosEdgeTp,
	PDL_ET_HomeMode.NegDirectionPosEdgeTp,
	PDL_ET_HomeMode.NegDirectionNegEdgeTp,
	PDL_ET_HomeMode.PosDirectionNegEdgeTp:
		fbHome.stTouchProbe := iq_stAxisModuleItf.stHome.stTouchProbe;

	PDL_ET_HomeMode.PosDirectionPosEdgeSensor,
	PDL_ET_HomeMode.NegDirectionPosEdgeSensor,
	PDL_ET_HomeMode.NegDirectionNegEdgeSensor,
	PDL_ET_HomeMode.PosDirectionNegEdgeSensor:
		fbHome.stSensor := iq_stAxisModuleItf.stHome.stSensor;

	PDL_ET_HomeMode.PosDirectionPosEdgeHWLimitPos,
	PDL_ET_HomeMode.NegDirectionPosEdgeHWLimitNeg,
	PDL_ET_HomeMode.NegDirectionNegEdgeHWLimitNeg,
	PDL_ET_HomeMode.PosDirectionNegEdgeHWLimitPos:
		fbHome.stLimitSwitch := iq_stAxisModuleItf.stHome.stLimitSwitch;

	PDL_ET_HomeMode.PosDirectionMaxTorque,
	PDL_ET_HomeMode.NegDirectionMaxTorque:
		fbHome.stTorque := iq_stAxisModuleItf.stHome.stTorque;

	PDL_ET_HomeMode.PosDirectionMaxForce,
	PDL_ET_HomeMode.NegDirectionMaxForce:
		fbHome.stForce:= iq_stAxisModuleItf.stHome.stForce;

	PDL_ET_HomeMode.MoveOnPosAbs:
		fbHome.stMoveOnPos := iq_stAxisModuleItf.stHome.stMoveonPos;

	PDL_ET_HomeMode.SetPosAxisPosition,
	PDL_ET_HomeMode.SetPosLogEncoderPosition,
	PDL_ET_HomeMode.SetPosAxisAndLogEncoderPosition,
	PDL_ET_HomeMode.RestorePosFromAxisEncoder,
	PDL_ET_HomeMode.RestorePosFromRetain:
		stFbHomeSetPosProperty.i_lrAbsEncOffset			:= iq_stAxisModuleItf.stHome.stSetPos.i_lrAbsEncOffset;
		stFbHomeSetPosProperty.i_lrEncoderPosition		:= iq_stAxisModuleItf.stHome.stSetPos.i_lrEncoderPosition;
		stFbHomeSetPosProperty.i_lrHomePosition			:= iq_stAxisModuleItf.stHome.stSetPos.i_lrHomePosition;
		stFbHomeSetPosProperty.i_lrRestoreWindow		:= iq_stAxisModuleItf.stHome.stSetPos.i_lrRestoreWindow;
		stFbHomeSetPosProperty.i_lrUserPeriod			:= iq_stAxisModuleItf.stHome.stSetPos.i_lrUserPeriod;
		stFbHomeSetPosProperty.iq_pstRestorePosRetain	:= iq_stAxisModuleItf.stHome.stSetPos.iq_pstRestorePosRetain;
		stFbHomeSetPosProperty.iq_lencAxis				:= iq_stAxisModuleItf.stMain.iq_lencEncoder;
		fbHome.stSetPos := stFbHomeSetPosProperty;

	PDL_ET_HomeMode.WriteAxisEncoder:
		fbHome.stWritePos := iq_stAxisModuleItf.stHome.stWritePos;
END_CASE

fbHome(	i_xEnable				:= xRefEnable AND (	   fbDriveEnable.q_xDriveEnabled
													OR fbHome.q_xDisableDrive
													OR xRefAxisEnableOld			(* xRefAxisEnableOld makes shure i_xEnable keeps true during reaktivation of axis after encoter writing *)
													OR iq_stAxisModuleItf.stHome.stSetPos.i_xKeepPowerDisabled),
		i_etMode				:= iq_stAxisModuleItf.stHome.i_etMode,
		i_ifDrive	 			:= iq_stAxisModuleItf.stMain.i_ifDrive,
		i_xHwLimitNeg			:= iq_stAxisModuleItf.stMain.i_xHwLimitNeg,
		i_xHwLimitPos			:= iq_stAxisModuleItf.stMain.i_xHwLimitPos,
		i_xStart				:= xRefStart,
		q_xActive				=> ,
		q_xReady				=> ,
		q_etDiag				=> etDiagBuffer,
		q_etDiagExt				=> etDiagExtBufferPDL,
		q_sMsg					=> sDiagMsgBuffer,
		q_xDisableDrive			=> ,
		q_xMotionInstructionActive	=> ,
		q_lrPosition			=> ,
		q_lrEncoderPosition		=> ,
		q_xHomeOk				=> );

DiagTestHoming(	iq_etDiag		:= fbHome.q_etDiag,
				iq_etDiagExt	:= fbHome.q_etDiagExt,
				iq_sMsg			:= fbHome.q_sMsg);

IF fbHome.i_xEnable THEN
	xRefAxisEnableOld := TRUE;
END_IF

IF fbHome.q_xHomeOk AND NOT xResetHomeOkActive THEN
	iq_stAxisModuleItf.stMain.q_xHomeOk := TRUE;
END_IF

IF fbHome.q_xReady AND NOT fbHome.i_xStart AND NOT fbHome.q_xHomeOk THEN
	iq_stAxisModuleItf.stMain.q_etState := AXM_ET_State.HomingWaitForStart;
ELSIF fbHome.q_xReady AND fbHome.i_xStart AND NOT fbHome.q_xHomeOk THEN
	iq_stAxisModuleItf.stMain.q_etState := AXM_ET_State.HomingExecuting;
ELSIF fbHome.q_xReady AND fbHome.q_xHomeOk AND NOT fbHome.q_xMotionInstructionActive THEN
	iq_stAxisModuleItf.stMain.q_etState := AXM_ET_State.HomingDone;
	xStartFlag := FALSE;
ELSE
	IF xRefEnable THEN
		iq_stAxisModuleItf.stMain.q_etState := AXM_ET_State.HomingInit;
	ELSE
		iq_stAxisModuleItf.stMain.q_etState := AXM_ET_State.HomingExit;
	END_IF
END_IF

IF NOT xRefEnable AND NOT fbHome.q_xActive THEN
	xRefActive := FALSE;
	xResetHomeOkActive := FALSE;
END_IF

IF xRefStart AND NOT xRefStartOld
		AND iq_stAxisModuleItf.stMain.i_ifDrive.etAxisState >= MOIN.ET_AxisState.Standstill
 		AND	iq_stAxisModuleItf.stMain.i_ifDrive.etAxisState <= MOIN.ET_AxisState.Stopping
		AND (  iq_stAxisModuleItf.stHome.i_etMode = PDL_ET_HomeMode.RestorePosFromAxisEncoder
			OR iq_stAxisModuleItf.stHome.i_etMode = PDL_ET_HomeMode.RestorePosFromRetain
			OR iq_stAxisModuleItf.stHome.i_etMode = PDL_ET_HomeMode.SetPosAxisAndLogEncoderPosition
			OR iq_stAxisModuleItf.stHome.i_etMode = PDL_ET_HomeMode.SetPosAxisPosition
			OR iq_stAxisModuleItf.stHome.i_etMode = PDL_ET_HomeMode.SetPosLogEncoderPosition )THEN

	ReadTrackingDeviation(	q_sLrealConversion => sLrealConversion);

	fbLoggerPoint.AddLogEntry (
			i_etLogLevel 	:= APL.ET_LogLevel.StatusMessage,
			i_etDiag		:= GD.ET_Diag.Ok,
			i_udiDiagExt	:= 0,
			i_sMessage		:= Standard.CONCAT('SetPos-Homing:  Axis-State >= Standstill; TrackingDeviation: ',sLrealConversion)
		);
END_IF
xRefStartOld := xRefStart;

(* ---- Homing_entry.act.st ---- *)
__METADATA__
{
  "v3Meta": {
    "objectGuid": "411e9c86-3a69-437b-80f4-8b885b1b2658",
    "objectTypeGuid": "8ac092e5-3128-4e26-9e7e-11016c6684f2",
    "embeddedObjectTypeGuids": [
      "3b83b776-fb25-43b8-99f2-3c507c9143fc"
    ],
    "properties": {},
    "subObjects": {}
  }
}

fbhome.RegisterLoggerPoint(	i_ifParent	:= fbLoggerPoint,
							i_sName		:= 'Homing',
							q_etDiag	=> ,
							q_etDiagExt => );

xRefActive := TRUE;
xRefAxisEnableOld := FALSE;

IF iq_stAxisModuleItf.stHome.i_etMode = PDL_ET_HomeMode.NegDirectionNegEdgeHWLimitNeg OR
	iq_stAxisModuleItf.stHome.i_etMode = PDL_ET_HomeMode.PosDirectionNegEdgeHWLimitPos THEN

	stExceptionModuleReaction2.etDiag 		:= GD.ET_Diag.ConfigurationFailed;
	stExceptionModuleReaction2.udiDiagExt 	:= AXM_ET_DiagExt.HomingModeNotSupported;
	stExceptionModuleReaction2.sMsg 		:= 'HomingMode LimitSwitch with NegEdge not supported. Use PosEdge inverted inputs';
	ReportException(iq_stException 	:= stExceptionModuleReaction2);

END_IF

(* ---- InactiveCmdExecution.meth.st ---- *)
{attribute 'conditionalshow_all_locals'}
METHOD INTERNAL InactiveCmdExecution
VAR_INPUT
END_VAR

(* Command execution if module is not active (q_xActive = FALSE) or currently deactivating (i_xEnable = FALSE, q_xActive is still TRUE) *)
IF iq_stStandardModuleItf.iq_diCmd <> 0 THEN
	IF(NOT iq_stStandardModuleItf.i_xEnable) THEN
		iq_stStandardModuleItf.iq_diCmd := 0; (* All commands are signaled executed if module is disabled *)
(*ELSE*)
	ELSIF(iq_stStandardModuleItf.iq_diCmd > 0) THEN (* New command *)
		(* Command execution during enable but module is not ready for commands yet ==> error *)
		//xExceptionCmdImpossibleState := TRUE;
		stExceptionCmdImpossibleState.udiDiagExt := AXM_ET_DiagExt.CmdImpossibleState;
		stExceptionCmdImpossibleState.sDiagExt := AXM_FC_EtDiagExtToString(i_etDiagExt := AXM_ET_DiagExt.CmdImpossibleState);
		stExceptionCmdImpossibleState.sMsg := SE_CTBX.FC_MultiConcat(	i_sString1 := 'Cmd impossible: ',
																	i_sString2 := AXM_FC_EtCmdToString(i_etCmd := ABS(iq_stStandardModuleItf.iq_diCMD)),
																	i_sString3 := '; State: ',
																	i_sString4 := AXM_FC_EtStateToString(i_etState := iq_stAxisModuleItf.stMain.q_etState));
		ReportException(iq_stException := stExceptionCmdImpossibleState);
		iq_stStandardModuleItf.iq_diCmd:= - ABS(iq_stStandardModuleItf.iq_diCmd);
	END_IF
END_IF
iq_stStandardModuleItf.q_xCmdActive := FALSE;
iq_stStandardModuleItf.q_xCmdDone := FALSE;
iq_stStandardModuleItf.q_diCmdActive := 0;
